{region 'Documentation'}
(*!
<summary>Selects explicit stimuli and expected outcomes; named constants identify every checkpoint.</summary>
*)
{endregion}
METHOD PRIVATE SelectStep : BOOL //! TRUE after selecting a supported script step and its literal expectations; FALSE reports an unknown step.
SelectStep := FALSE;
FRisingFindingExpected := FALSE;
FFallingFindingExpected := FALSE;
FDelayedRisingFindingExpected := FALSE;
FDelayedFallingFindingExpected := FALSE;
CASE FStep OF
    StepInitialBoundReset:
        FTrace := TraceResetHistory;
        FSample := TRUE;
        FSubjectEnable := TRUE;
        FResetSubjects := TRUE;
        FExpectedResult := E_Result.NotEvaluated;
        FExpectedDelayedResult := E_Result.NotEvaluated;
        FExpectedObservation := FALSE;
        FExpectedDelayedObservation := FALSE;
        FExpectedEvaluation := FALSE;
        FExpectedDelayedEvaluation := FALSE;
    StepFirstHighSample:
        FTrace := TraceFirstObservation;
        FSample := TRUE;
        FSubjectEnable := TRUE;
        FResetSubjects := FALSE;
        FExpectedResult := E_Result.NotEvaluated;
        FExpectedDelayedResult := E_Result.NotEvaluated;
        FExpectedObservation := TRUE;
        FExpectedDelayedObservation := FALSE;
        FExpectedEvaluation := FALSE;
        FExpectedDelayedEvaluation := FALSE;
    StepSameHighSample:
        FTrace := TraceFirstObservation;
        FSample := TRUE;
        FSubjectEnable := TRUE;
        FResetSubjects := FALSE;
        FExpectedResult := E_Result.Passed;
        FExpectedDelayedResult := E_Result.NotEvaluated;
        FExpectedObservation := TRUE;
        FExpectedDelayedObservation := TRUE;
        FExpectedEvaluation := TRUE;
        FExpectedDelayedEvaluation := FALSE;
    StepOppositeEdgeAllowed:
        FTrace := TraceFirstObservation;
        FSample := FALSE;
        FSubjectEnable := TRUE;
        FResetSubjects := FALSE;
        FExpectedResult := E_Result.Passed;
        FExpectedDelayedResult := E_Result.Passed;
        FExpectedObservation := TRUE;
        FExpectedDelayedObservation := TRUE;
        FExpectedEvaluation := TRUE;
        FExpectedDelayedEvaluation := TRUE;
    StepForbiddenEdge:
        FTrace := TraceHeldFailure;
        FSample := TRUE;
        FSubjectEnable := TRUE;
        FResetSubjects := FALSE;
        FExpectedResult := E_Result.Failed;
        FExpectedDelayedResult := E_Result.Failed;
        FExpectedObservation := TRUE;
        FExpectedDelayedObservation := TRUE;
        FExpectedEvaluation := TRUE;
        FExpectedDelayedEvaluation := TRUE;
        FRisingFindingExpected := TRUE;
        FFallingFindingExpected := TRUE;
        FDelayedRisingFindingExpected := TRUE;
        FDelayedFallingFindingExpected := TRUE;
    StepRepeatedFailure:
        FTrace := TraceHeldFailure;
        FSample := TRUE;
        FSubjectEnable := TRUE;
        FResetSubjects := FALSE;
        FExpectedResult := E_Result.Failed;
        FExpectedDelayedResult := E_Result.Failed;
        FExpectedObservation := TRUE;
        FExpectedDelayedObservation := TRUE;
        FExpectedEvaluation := TRUE;
        FExpectedDelayedEvaluation := TRUE;
    StepResetBeforeGap:
        FTrace := TraceResetHistory;
        FSample := FALSE;
        FSubjectEnable := TRUE;
        FResetSubjects := TRUE;
        FExpectedResult := E_Result.NotEvaluated;
        FExpectedDelayedResult := E_Result.NotEvaluated;
        FExpectedObservation := FALSE;
        FExpectedDelayedObservation := FALSE;
        FExpectedEvaluation := FALSE;
        FExpectedDelayedEvaluation := FALSE;
    StepBaselineBeforeGap:
        FTrace := TraceDisabledHistory;
        FSample := FALSE;
        FSubjectEnable := TRUE;
        FResetSubjects := FALSE;
        FExpectedResult := E_Result.NotEvaluated;
        FExpectedDelayedResult := E_Result.NotEvaluated;
        FExpectedObservation := TRUE;
        FExpectedDelayedObservation := FALSE;
        FExpectedEvaluation := FALSE;
        FExpectedDelayedEvaluation := FALSE;
    StepDisabledChange:
        FTrace := TraceDisabledHistory;
        FSample := TRUE;
        FSubjectEnable := FALSE;
        FResetSubjects := FALSE;
        FExpectedResult := E_Result.NotEvaluated;
        FExpectedDelayedResult := E_Result.NotEvaluated;
        FExpectedObservation := FALSE;
        FExpectedDelayedObservation := FALSE;
        FExpectedEvaluation := FALSE;
        FExpectedDelayedEvaluation := FALSE;
    StepFirstAfterGap:
        FTrace := TraceDisabledHistory;
        FSample := TRUE;
        FSubjectEnable := TRUE;
        FResetSubjects := FALSE;
        FExpectedResult := E_Result.NotEvaluated;
        FExpectedDelayedResult := E_Result.NotEvaluated;
        FExpectedObservation := TRUE;
        FExpectedDelayedObservation := FALSE;
        FExpectedEvaluation := FALSE;
        FExpectedDelayedEvaluation := FALSE;
    StepSecondAfterGap:
        FTrace := TraceDisabledHistory;
        FSample := TRUE;
        FSubjectEnable := TRUE;
        FResetSubjects := FALSE;
        FExpectedResult := E_Result.Passed;
        FExpectedDelayedResult := E_Result.NotEvaluated;
        FExpectedObservation := TRUE;
        FExpectedDelayedObservation := TRUE;
        FExpectedEvaluation := TRUE;
        FExpectedDelayedEvaluation := FALSE;
    StepAllowedAfterGap:
        FTrace := TraceDisabledHistory;
        FSample := FALSE;
        FSubjectEnable := TRUE;
        FResetSubjects := FALSE;
        FExpectedResult := E_Result.Passed;
        FExpectedDelayedResult := E_Result.Passed;
        FExpectedObservation := TRUE;
        FExpectedDelayedObservation := TRUE;
        FExpectedEvaluation := TRUE;
        FExpectedDelayedEvaluation := TRUE;
    StepForbiddenAfterGap:
        FTrace := TraceDisabledHistory;
        FSample := TRUE;
        FSubjectEnable := TRUE;
        FResetSubjects := FALSE;
        FExpectedResult := E_Result.Failed;
        FExpectedDelayedResult := E_Result.Failed;
        FExpectedObservation := TRUE;
        FExpectedDelayedObservation := TRUE;
        FExpectedEvaluation := TRUE;
        FExpectedDelayedEvaluation := TRUE;
        FRisingFindingExpected := TRUE;
        FFallingFindingExpected := TRUE;
        FDelayedRisingFindingExpected := TRUE;
        FDelayedFallingFindingExpected := TRUE;
    StepResetBeforeDelay:
        FTrace := TraceResetHistory;
        FSample := FALSE;
        FSubjectEnable := TRUE;
        FResetSubjects := TRUE;
        FExpectedResult := E_Result.NotEvaluated;
        FExpectedDelayedResult := E_Result.NotEvaluated;
        FExpectedObservation := FALSE;
        FExpectedDelayedObservation := FALSE;
        FExpectedEvaluation := FALSE;
        FExpectedDelayedEvaluation := FALSE;
    StepSkippedFirstBaseline:
        FTrace := TraceDelayedObservation;
        FSample := FALSE;
        FSubjectEnable := TRUE;
        FResetSubjects := FALSE;
        FExpectedResult := E_Result.NotEvaluated;
        FExpectedDelayedResult := E_Result.NotEvaluated;
        FExpectedObservation := TRUE;
        FExpectedDelayedObservation := FALSE;
        FExpectedEvaluation := FALSE;
        FExpectedDelayedEvaluation := FALSE;
    StepEdgeBeforeDelayedBaseline:
        FTrace := TraceDelayedObservation;
        FSample := TRUE;
        FSubjectEnable := TRUE;
        FResetSubjects := FALSE;
        FExpectedResult := E_Result.Failed;
        FExpectedDelayedResult := E_Result.NotEvaluated;
        FExpectedObservation := TRUE;
        FExpectedDelayedObservation := TRUE;
        FExpectedEvaluation := TRUE;
        FExpectedDelayedEvaluation := FALSE;
        FRisingFindingExpected := TRUE;
        FFallingFindingExpected := TRUE;
    StepStableDelayedBaseline:
        FTrace := TraceDelayedObservation;
        FSample := TRUE;
        FSubjectEnable := TRUE;
        FResetSubjects := FALSE;
        FExpectedResult := E_Result.Failed;
        FExpectedDelayedResult := E_Result.Passed;
        FExpectedObservation := TRUE;
        FExpectedDelayedObservation := TRUE;
        FExpectedEvaluation := TRUE;
        FExpectedDelayedEvaluation := TRUE;
ELSE
    Error(Message := 'Unknown observation trace step.');
    RETURN;
END_CASE;
SelectStep := TRUE;
END_METHOD

END_FUNCTION_BLOCK

// ---- SelfTests/TestCases/TestSuite_AssertionObservation/Test_AssertionEdgeCount.TcPOU
{region 'Documentation'}
(*!
<summary>Checks accumulated rising/falling counts and independent evaluation timing.</summary>
<description>
Both directions run with normal and delayed first observation. Counts survive disabled intervals, but transitions across a gap do not count. Combined observation/evaluation includes the current edge; Evaluate alone observes no edge. Literal counts test the shared algorithm without repeating the comparison operator matrix.
ProcessTests executes one named step per PLC cycle. ProcessAssertions checks that
step before the next call advances it. Every trace has its own outer Assertion;
FirstFailedStep retains the first mismatching checkpoint for online diagnosis.
Expected findings are captured locally and checked before the next step clears
that capture. Subjects are deliberately not called between scripted steps.
</description>
*)
{endregion}
FUNCTION_BLOCK Test_AssertionEdgeCount EXTENDS TestCaseBase
VAR
    FRising : AssertRisingEdgeCntEqual;
    FFalling : AssertFallingEdgeCntEqual;
    FDelayedRising : AssertRisingEdgeCntEqual;
    FDelayedFalling : AssertFallingEdgeCntEqual;
    FCapture : EventBuffer;
    FEvents : ARRAY[1..CaptureLength] OF ST_Event;
    FCaptureFifo : ST_FifoStatus;
    FCaptureStatus : ST_EventBufferStatus;
    FSetupValid : BOOL;
    FStep : UINT;
    FTrace : UINT;
    FFirstFailedStep : UINT;
    FChecked : BOOL;
    FObservationReady : BOOL;
    FStepMatches : BOOL;
    FResultsMatch : BOOL;
    FActivityMatches : BOOL;
    FFindingsMatch : BOOL;
    FCountsMatch : BOOL;
    FSample : BOOL;
    FSubjectEnable : BOOL;
    FSubjectEvaluate : BOOL;
    FResetSubjects : BOOL;
    FExpectedResult : E_Result;
    FExpectedDelayedResult : E_Result;
    FExpectedObservation : BOOL;
    FExpectedDelayedObservation : BOOL;
    FExpectedEvaluation : BOOL;
    FExpectedDelayedEvaluation : BOOL;
    FCountTarget : UINT;
    FExpectedCount : UINT;
    FRisingFindingExpected : BOOL;
    FFallingFindingExpected : BOOL;
    FDelayedRisingFindingExpected : BOOL;
    FDelayedFallingFindingExpected : BOOL;
END_VAR
VAR
    FResetHistory : AssertTrue;
    FCounting : AssertTrue;
    FDisabledHistory : AssertTrue;
    FEvaluationTiming : AssertTrue;
    FWrongCount : AssertTrue;
END_VAR
VAR CONSTANT
    CaptureLength : UINT := 8;
    StepInitialBoundReset : UINT := 1;
    StepFirstBaseline : UINT := 2;
    StepRepeatedBaseline : UINT := 3;
    StepFirstEdge : UINT := 4;
    StepHeldSignal : UINT := 5;
    StepOppositeEdge : UINT := 6;
    StepSecondEdge : UINT := 7;
    StepDisabledChange : UINT := 8;
    StepFirstAfterGap : UINT := 9;
    StepSecondAfterGap : UINT := 10;
    StepOppositeAfterGap : UINT := 11;
    StepThirdEdge : UINT := 12;
    StepEvaluateOnly : UINT := 13;
    StepBaselineBeforeCombined : UINT := 14;
    StepLowBeforeCombined : UINT := 15;
    StepCountBeforeEvaluate : UINT := 16;
    StepResetAfterPass : UINT := 17;
    StepEvaluateOnFirstEnable : UINT := 18;
    StepNewLowBaseline : UINT := 19;
    StepWrongCountFinding : UINT := 20;
    StepWrongCountHeld : UINT := 21;
    StepResetAfterFailure : UINT := 22;
    LastStep : UINT := StepResetAfterFailure;
    TraceResetHistory : UINT := 1;
    TraceCounting : UINT := 2;
    TraceDisabledHistory : UINT := 3;
    TraceEvaluationTiming : UINT := 4;
    TraceWrongCount : UINT := 5;
END_VAR

SUPER^();

{region 'Documentation'}
(*!
<summary>Collects the outer trace checks, never subject results.</summary>
*)
{endregion}
METHOD PROTECTED AggregateResults
VAR_INPUT
    Aggregator : I_ResultAggregator; //! Borrowed result sink owned by the outer Test Case; add this test's checking Assertions without resetting or retaining the sink.
END_VAR
Aggregator.AddProvider(Provider := FResetHistory);
Aggregator.AddProvider(Provider := FCounting);
Aggregator.AddProvider(Provider := FDisabledHistory);
Aggregator.AddProvider(Provider := FEvaluationTiming);
Aggregator.AddProvider(Provider := FWrongCount);
END_METHOD

{region 'Documentation'}
(*!
<summary>Calls each real production subject once with this step's bound inputs.</summary>
*)
{endregion}
METHOD PRIVATE CallSubjects
FRising(Enable := FSubjectEnable,
    Evaluate := FSubjectEvaluate,
    State := E_State.Running,
    IN := FSample,
    Expected := FCountTarget);
FFalling(Enable := FSubjectEnable,
    Evaluate := FSubjectEvaluate,
    State := E_State.Running,
    IN := NOT FSample,
    Expected := FCountTarget);
FDelayedRising(Enable := FSubjectEnable,
    Evaluate := FSubjectEvaluate,
    State := E_State.Running,
    IN := FSample,
    Expected := FCountTarget);
FDelayedFalling(Enable := FSubjectEnable,
    Evaluate := FSubjectEvaluate,
    State := E_State.Running,
    IN := NOT FSample,
    Expected := FCountTarget);
END_METHOD

{region 'Documentation'}
(*!
<summary>Checks per-step finding order, identity and count without retaining old events.</summary>
*)
{endregion}
METHOD PRIVATE CheckFindings
VAR
    Index : UINT;
    FindingMatches : BOOL;
END_VAR
Index := 1;
FFindingsMatch := TRUE;
IF FRisingFindingExpected THEN
    FindingMatches := IsFindingValid(Index := Index,
        ExpectedName := FRising.Name);
    FFindingsMatch := FFindingsMatch AND FindingMatches;
    Index := Index + 1;
END_IF;
IF FFallingFindingExpected THEN
    FindingMatches := IsFindingValid(Index := Index,
        ExpectedName := FFalling.Name);
    FFindingsMatch := FFindingsMatch AND FindingMatches;
    Index := Index + 1;
END_IF;
IF FDelayedRisingFindingExpected THEN
    FindingMatches := IsFindingValid(Index := Index,
        ExpectedName := FDelayedRising.Name);
    FFindingsMatch := FFindingsMatch AND FindingMatches;
    Index := Index + 1;
END_IF;
IF FDelayedFallingFindingExpected THEN
    FindingMatches := IsFindingValid(Index := Index,
        ExpectedName := FDelayedFalling.Name);
    FFindingsMatch := FFindingsMatch AND FindingMatches;
    Index := Index + 1;
END_IF;
FFindingsMatch := FFindingsMatch
    AND (FCaptureStatus.SequenceId = UINT_TO_UDINT(Index - 1))
    AND (FCaptureStatus.LostEventCount = 0);
END_METHOD

{region 'Documentation'}
(*!
<summary>Rejects incomplete local capture, subject or checking-Assertion setup.</summary>
*)
{endregion}
METHOD PROTECTED CheckInitialization : BOOL //! TRUE when the inherited initialization check and this concrete fixture check both accept the setup.
CheckInitialization := SUPER^.CheckInitialization();
IF NOT CheckInitialization THEN
    RETURN;
END_IF;

CheckInitialization := FSetupValid
    AND FResetHistory.IsInitialized
    AND FCounting.IsInitialized
    AND FDisabledHistory.IsInitialized
    AND FEvaluationTiming.IsInitialized
    AND FWrongCount.IsInitialized;
IF NOT CheckInitialization THEN
    EventPublisher.PublishEvent(Event := CreateFrameworkEvent(Name := Name,
        ResourceName := '',
        State := State,
        Severity := E_EventSeverity.Error,
        Message := 'Observation selftest setup failed.'));
END_IF;
END_METHOD

{region 'Documentation'}
(*!
<summary>Compares public results and activity gates against literal step expectations.</summary>
*)
{endregion}
METHOD PRIVATE CheckResults
FResultsMatch := (FRising.Result = FExpectedResult)
    AND (FFalling.Result = FExpectedResult)
    AND (FDelayedRising.Result = FExpectedDelayedResult)
    AND (FDelayedFalling.Result = FExpectedDelayedResult);
FActivityMatches := (FRising.Enabled = FSubjectEnable)
    AND (FRising.ObservationActive = FExpectedObservation)
    AND (FRising.EvaluationActive = FExpectedEvaluation)
    AND (FFalling.Enabled = FSubjectEnable)
    AND (FFalling.ObservationActive = FExpectedObservation)
    AND (FFalling.EvaluationActive = FExpectedEvaluation)
    AND (FDelayedRising.Enabled = FSubjectEnable)
    AND (FDelayedRising.ObservationActive = FExpectedDelayedObservation)
    AND (FDelayedRising.EvaluationActive = FExpectedDelayedEvaluation)
    AND (FDelayedFalling.Enabled = FSubjectEnable)
    AND (FDelayedFalling.ObservationActive = FExpectedDelayedObservation)
    AND (FDelayedFalling.EvaluationActive = FExpectedDelayedEvaluation);
FCountsMatch := (FRising.EdgeCount = FExpectedCount)
    AND (FFalling.EdgeCount = FExpectedCount)
    AND (FDelayedRising.EdgeCount = FExpectedCount)
    AND (FDelayedFalling.EdgeCount = FExpectedCount);
END_METHOD

{region 'Documentation'}
(*!
<summary>Binds isolated subjects and initializes the outer trace Assertions.</summary>
*)
{endregion}
METHOD PROTECTED Configure
VAR
    Initialized : BOOL;
END_VAR
FPreparationStateCount := 0;
FTestStateCount := 1;
FResetHistory.Initialize(Parent := THIS^,
    AssertionName := 'ResetHistory');
FCounting.Initialize(Parent := THIS^,
    AssertionName := 'Counting');
FDisabledHistory.Initialize(Parent := THIS^,
    AssertionName := 'DisabledHistory');
FEvaluationTiming.Initialize(Parent := THIS^,
    AssertionName := 'EvaluationTiming');
FWrongCount.Initialize(Parent := THIS^,
    AssertionName := 'WrongCount');
FSetupValid := FCapture.Initialize(Buffer := FEvents,
    FifoControl := FCaptureFifo,
    Status := FCaptureStatus);
FRising.BindPublisher(Publisher := FCapture);
Initialized := FRising.Initialize(Parent := THIS^,
    AssertionName := 'Rising',
    ObserveFirstCycle := TRUE);
FSetupValid := FSetupValid AND Initialized;
FFalling.BindPublisher(Publisher := FCapture);
Initialized := FFalling.Initialize(Parent := THIS^,
    AssertionName := 'Falling',
    ObserveFirstCycle := TRUE);
FSetupValid := FSetupValid AND Initialized;
FDelayedRising.BindPublisher(Publisher := FCapture);
Initialized := FDelayedRising.Initialize(Parent := THIS^,
    AssertionName := 'DelayedRising',
    ObserveFirstCycle := FALSE);
FSetupValid := FSetupValid AND Initialized;
FDelayedFalling.BindPublisher(Publisher := FCapture);
Initialized := FDelayedFalling.Initialize(Parent := THIS^,
    AssertionName := 'DelayedFalling',
    ObserveFirstCycle := FALSE);
FSetupValid := FSetupValid AND Initialized;
END_METHOD

{region 'Documentation'}
(*!
<summary>Checks one expected local Failed finding; index is bounded by four subjects.</summary>
*)
{endregion}
METHOD PRIVATE IsFindingValid : BOOL //! TRUE when the selected captured finding satisfies the scenario metadata and diagnostic checks.
VAR_INPUT
    Index : UINT; //! One-based index in the retained isolated event capture.
    ExpectedName : STRING(GVL_Constants.NameLength); //! Independently authored Assertion name expected in the selected finding.
END_VAR
IsFindingValid := (FEvents[Index].SequenceId = UINT_TO_UDINT(Index))
    AND (FEvents[Index].Name = ExpectedName)
    AND (FEvents[Index].OwnerScope = E_OwnerScope.Assertion)
    AND (FEvents[Index].EventType = E_EventType.Result)
    AND (FEvents[Index].State = E_State.Running)
    AND (FEvents[Index].Result = E_Result.Failed)
    AND (FEvents[Index].Message <> '');
END_METHOD

{region 'Documentation'}
(*!
<summary>Completes abort; the trace owns no asynchronous resource.</summary>
*)
{endregion}
METHOD PROTECTED ProcessAbort
VAR_INPUT
    Enable : BOOL; //! Phase permission supplied by the owning Test Case; FALSE does not authorize progression, while observation may continue.
END_VAR
IF Enable THEN
    CompleteAbort();
END_IF;
END_METHOD

{region 'Documentation'}
(*!
<summary>Latches the current trace checkpoint before allowing progression.</summary>
*)
{endregion}
METHOD PROTECTED ProcessAssertions
VAR_INPUT
    Enable : BOOL; //! Phase permission supplied by the owning Test Case; FALSE does not authorize progression, while observation may continue.
END_VAR
VAR
    Check : BOOL;
END_VAR
Check := Enable AND FObservationReady;
FResetHistory(Enable := Check AND (FTrace = TraceResetHistory),
    State := State,
    IN := FStepMatches);
FCounting(Enable := Check AND (FTrace = TraceCounting),
    State := State,
    IN := FStepMatches);
FDisabledHistory(Enable := Check AND (FTrace = TraceDisabledHistory),
    State := State,
    IN := FStepMatches);
FEvaluationTiming(Enable := Check AND (FTrace = TraceEvaluationTiming),
    State := State,
    IN := FStepMatches);
FWrongCount(Enable := Check AND (FTrace = TraceWrongCount),
    State := State,
    IN := FStepMatches);
IF Check THEN
    FChecked := TRUE;
END_IF;
END_METHOD

{region 'Documentation'}
(*!
<summary>No Preparation phase is required.</summary>
*)
{endregion}
METHOD PROTECTED ProcessPreparations
VAR_INPUT
    // SA0033: Required hook; this test has no Preparation phase.
    {attribute 'analysis' := '-33'}
    Enable : BOOL; //! Phase permission supplied by the owning Test Case; FALSE does not authorize progression, while observation may continue.
END_VAR
END_METHOD

{region 'Documentation'}
(*!
<summary>Restarts the trace; subjects consume their reset only with bound inputs.</summary>
*)
{endregion}
METHOD PROTECTED ProcessReset
FStep := StepInitialBoundReset;
FTrace := 0;
FFirstFailedStep := 0;
FChecked := FALSE;
FObservationReady := FALSE;
FStepMatches := TRUE;
FResultsMatch := TRUE;
FActivityMatches := TRUE;
FFindingsMatch := TRUE;
FCountsMatch := TRUE;
FCapture.Reset();
ResetSubjects();
FResetHistory.Reset();
FCounting.Reset();
FDisabledHistory.Reset();
FEvaluationTiming.Reset();
FWrongCount.Reset();
CompleteReset();
END_METHOD

{region 'Documentation'}
(*!
<summary>Executes one named step per active cycle, after the previous check was latched.</summary>
*)
{endregion}
METHOD PROTECTED ProcessTests
VAR_INPUT
    Enable : BOOL; //! Phase permission supplied by the owning Test Case; FALSE does not authorize progression, while observation may continue.
END_VAR
IF NOT Enable THEN
    RETURN;
END_IF;

IF FChecked THEN
    FChecked := FALSE;
    FObservationReady := FALSE;
    IF FStep = LastStep THEN
        CompleteTests();
        RETURN;
    END_IF;
    FStep := FStep + 1;
END_IF;

IF NOT SelectStep() THEN
    RETURN;
END_IF;
FCapture.Reset();
IF FResetSubjects THEN
    ResetSubjects();
END_IF;
CallSubjects();
CheckResults();
CheckFindings();
FStepMatches := FResultsMatch AND FActivityMatches AND FFindingsMatch AND FCountsMatch;
IF NOT FStepMatches AND (FFirstFailedStep = 0) THEN
    FFirstFailedStep := FStep;
END_IF;
FObservationReady := TRUE;
END_METHOD

{region 'Documentation'}
(*!
<summary>Queues reset without accessing typed cyclic inputs.</summary>
*)
{endregion}
METHOD PRIVATE ResetSubjects
FRising.Reset();
FFalling.Reset();
FDelayedRising.Reset();
FDelayedFalling.Reset();
END_METHOD

{region 'Documentation'}
(*!
<summary>Selects explicit stimuli and expected outcomes; named constants identify every checkpoint.</summary>
*)
{endregion}
METHOD PRIVATE SelectStep : BOOL //! TRUE after selecting a supported script step and its literal expectations; FALSE reports an unknown step.
SelectStep := FALSE;
FRisingFindingExpected := FALSE;
FFallingFindingExpected := FALSE;
FDelayedRisingFindingExpected := FALSE;
FDelayedFallingFindingExpected := FALSE;
CASE FStep OF
    StepInitialBoundReset:
        FTrace := TraceResetHistory;
        FSample := FALSE;
        FSubjectEnable := TRUE;
        FSubjectEvaluate := FALSE;
        FResetSubjects := TRUE;
        FExpectedResult := E_Result.NotEvaluated;
        FExpectedDelayedResult := E_Result.NotEvaluated;
        FExpectedObservation := FALSE;
        FExpectedDelayedObservation := FALSE;
        FExpectedEvaluation := FALSE;
        FExpectedDelayedEvaluation := FALSE;
        FExpectedCount := 0;
        FCountTarget := 0;
    StepFirstBaseline:
        FTrace := TraceCounting;
        FSample := FALSE;
        FSubjectEnable := TRUE;
        FSubjectEvaluate := FALSE;
        FResetSubjects := FALSE;
        FExpectedResult := E_Result.NotEvaluated;
        FExpectedDelayedResult := E_Result.NotEvaluated;
        FExpectedObservation := TRUE;
        FExpectedDelayedObservation := FALSE;
        FExpectedEvaluation := FALSE;
        FExpectedDelayedEvaluation := FALSE;
        FExpectedCount := 0;
        FCountTarget := 0;
    StepRepeatedBaseline:
        FTrace := TraceCounting;
        FSample := FALSE;
        FSubjectEnable := TRUE;
        FSubjectEvaluate := FALSE;
        FResetSubjects := FALSE;
        FExpectedResult := E_Result.NotEvaluated;
        FExpectedDelayedResult := E_Result.NotEvaluated;
        FExpectedObservation := TRUE;
        FExpectedDelayedObservation := TRUE;
        FExpectedEvaluation := FALSE;
        FExpectedDelayedEvaluation := FALSE;
        FExpectedCount := 0;
        FCountTarget := 0;
    StepFirstEdge:
        FTrace := TraceCounting;
        FSample := TRUE;
        FSubjectEnable := TRUE;
        FSubjectEvaluate := FALSE;
        FResetSubjects := FALSE;
        FExpectedResult := E_Result.NotEvaluated;
        FExpectedDelayedResult := E_Result.NotEvaluated;
        FExpectedObservation := TRUE;
        FExpectedDelayedObservation := TRUE;
        FExpectedEvaluation := FALSE;
        FExpectedDelayedEvaluation := FALSE;
        FExpectedCount := 1;
        FCountTarget := 0;
    StepHeldSignal:
        FTrace := TraceCounting;
        FSample := TRUE;
        FSubjectEnable := TRUE;
        FSubjectEvaluate := FALSE;
        FResetSubjects := FALSE;
        FExpectedResult := E_Result.NotEvaluated;
        FExpectedDelayedResult := E_Result.NotEvaluated;
        FExpectedObservation := TRUE;
        FExpectedDelayedObservation := TRUE;
        FExpectedEvaluation := FALSE;
        FExpectedDelayedEvaluation := FALSE;
        FExpectedCount := 1;
        FCountTarget := 0;
    StepOppositeEdge:
        FTrace := TraceCounting;
        FSample := FALSE;
        FSubjectEnable := TRUE;
        FSubjectEvaluate := FALSE;
        FResetSubjects := FALSE;
        FExpectedResult := E_Result.NotEvaluated;
        FExpectedDelayedResult := E_Result.NotEvaluated;
        FExpectedObservation := TRUE;
        FExpectedDelayedObservation := TRUE;
        FExpectedEvaluation := FALSE;
        FExpectedDelayedEvaluation := FALSE;
        FExpectedCount := 1;
        FCountTarget := 0;
    StepSecondEdge:
        FTrace := TraceCounting;
        FSample := TRUE;
        FSubjectEnable := TRUE;
        FSubjectEvaluate := FALSE;
        FResetSubjects := FALSE;
        FExpectedResult := E_Result.NotEvaluated;
        FExpectedDelayedResult := E_Result.NotEvaluated;
        FExpectedObservation := TRUE;
        FExpectedDelayedObservation := TRUE;
        FExpectedEvaluation := FALSE;
        FExpectedDelayedEvaluation := FALSE;
        FExpectedCount := 2;
        FCountTarget := 0;
    StepDisabledChange:
        FTrace := TraceDisabledHistory;
        FSample := FALSE;
        FSubjectEnable := FALSE;
        FSubjectEvaluate := FALSE;
        FResetSubjects := FALSE;
        FExpectedResult := E_Result.NotEvaluated;
        FExpectedDelayedResult := E_Result.NotEvaluated;
        FExpectedObservation := FALSE;
        FExpectedDelayedObservation := FALSE;
        FExpectedEvaluation := FALSE;
        FExpectedDelayedEvaluation := FALSE;
        FExpectedCount := 2;
        FCountTarget := 0;
    StepFirstAfterGap:
        FTrace := TraceDisabledHistory;
        FSample := TRUE;
        FSubjectEnable := TRUE;
        FSubjectEvaluate := FALSE;
        FResetSubjects := FALSE;
        FExpectedResult := E_Result.NotEvaluated;
        FExpectedDelayedResult := E_Result.NotEvaluated;
        FExpectedObservation := TRUE;
        FExpectedDelayedObservation := FALSE;
        FExpectedEvaluation := FALSE;
        FExpectedDelayedEvaluation := FALSE;
        FExpectedCount := 2;
        FCountTarget := 0;
    StepSecondAfterGap:
        FTrace := TraceDisabledHistory;
        FSample := TRUE;
        FSubjectEnable := TRUE;
        FSubjectEvaluate := FALSE;
        FResetSubjects := FALSE;
        FExpectedResult := E_Result.NotEvaluated;
        FExpectedDelayedResult := E_Result.NotEvaluated;
        FExpectedObservation := TRUE;
        FExpectedDelayedObservation := TRUE;
        FExpectedEvaluation := FALSE;
        FExpectedDelayedEvaluation := FALSE;
        FExpectedCount := 2;
        FCountTarget := 0;
    StepOppositeAfterGap:
        FTrace := TraceDisabledHistory;
        FSample := FALSE;
        FSubjectEnable := TRUE;
        FSubjectEvaluate := FALSE;
        FResetSubjects := FALSE;
        FExpectedResult := E_Result.NotEvaluated;
        FExpectedDelayedResult := E_Result.NotEvaluated;
        FExpectedObservation := TRUE;
        FExpectedDelayedObservation := TRUE;
        FExpectedEvaluation := FALSE;
        FExpectedDelayedEvaluation := FALSE;
        FExpectedCount := 2;
        FCountTarget := 0;
    StepThirdEdge:
        FTrace := TraceDisabledHistory;
        FSample := TRUE;
        FSubjectEnable := TRUE;
        FSubjectEvaluate := FALSE;
        FResetSubjects := FALSE;
        FExpectedResult := E_Result.NotEvaluated;
        FExpectedDelayedResult := E_Result.NotEvaluated;
        FExpectedObservation := TRUE;
        FExpectedDelayedObservation := TRUE;
        FExpectedEvaluation := FALSE;
        FExpectedDelayedEvaluation := FALSE;
        FExpectedCount := 3;
        FCountTarget := 0;
    StepEvaluateOnly:
        FTrace := TraceEvaluationTiming;
        FSample := FALSE;
        FSubjectEnable := FALSE;
        FSubjectEvaluate := TRUE;
        FResetSubjects := FALSE;
        FExpectedResult := E_Result.Passed;
        FExpectedDelayedResult := E_Result.Passed;
        FExpectedObservation := FALSE;
        FExpectedDelayedObservation := FALSE;
        FExpectedEvaluation := TRUE;
        FExpectedDelayedEvaluation := TRUE;
        FExpectedCount := 3;
        FCountTarget := 3;
    StepBaselineBeforeCombined:
        FTrace := TraceEvaluationTiming;
        FSample := TRUE;
        FSubjectEnable := TRUE;
        FSubjectEvaluate := FALSE;
        FResetSubjects := FALSE;
        FExpectedResult := E_Result.Passed;
        FExpectedDelayedResult := E_Result.Passed;
        FExpectedObservation := TRUE;
        FExpectedDelayedObservation := FALSE;
        FExpectedEvaluation := FALSE;
        FExpectedDelayedEvaluation := FALSE;
        FExpectedCount := 3;
        FCountTarget := 0;
    StepLowBeforeCombined:
        FTrace := TraceEvaluationTiming;
        FSample := FALSE;
        FSubjectEnable := TRUE;
        FSubjectEvaluate := FALSE;
        FResetSubjects := FALSE;
        FExpectedResult := E_Result.Passed;
        FExpectedDelayedResult := E_Result.Passed;
        FExpectedObservation := TRUE;
        FExpectedDelayedObservation := TRUE;
        FExpectedEvaluation := FALSE;
        FExpectedDelayedEvaluation := FALSE;
        FExpectedCount := 3;
        FCountTarget := 0;
    StepCountBeforeEvaluate:
        FTrace := TraceEvaluationTiming;
        FSample := TRUE;
        FSubjectEnable := TRUE;
        FSubjectEvaluate := TRUE;
        FResetSubjects := FALSE;
        FExpectedResult := E_Result.Passed;
        FExpectedDelayedResult := E_Result.Passed;
        FExpectedObservation := TRUE;
        FExpectedDelayedObservation := TRUE;
        FExpectedEvaluation := TRUE;
        FExpectedDelayedEvaluation := TRUE;
        FExpectedCount := 4;
        FCountTarget := 4;
    StepResetAfterPass:
        FTrace := TraceResetHistory;
        FSample := TRUE;
        FSubjectEnable := TRUE;
        FSubjectEvaluate := TRUE;
        FResetSubjects := TRUE;
        FExpectedResult := E_Result.NotEvaluated;
        FExpectedDelayedResult := E_Result.NotEvaluated;
        FExpectedObservation := FALSE;
        FExpectedDelayedObservation := FALSE;
        FExpectedEvaluation := FALSE;
        FExpectedDelayedEvaluation := FALSE;
        FExpectedCount := 0;
        FCountTarget := 0;
    StepEvaluateOnFirstEnable:
        FTrace := TraceEvaluationTiming;
        FSample := TRUE;
        FSubjectEnable := TRUE;
        FSubjectEvaluate := TRUE;
        FResetSubjects := FALSE;
        FExpectedResult := E_Result.Passed;
        FExpectedDelayedResult := E_Result.Passed;
        FExpectedObservation := TRUE;
        FExpectedDelayedObservation := FALSE;
        FExpectedEvaluation := TRUE;
        FExpectedDelayedEvaluation := TRUE;
        FExpectedCount := 0;
        FCountTarget := 0;
    StepNewLowBaseline:
        FTrace := TraceWrongCount;
        FSample := FALSE;
        FSubjectEnable := TRUE;
        FSubjectEvaluate := FALSE;
        FResetSubjects := FALSE;
        FExpectedResult := E_Result.Passed;
        FExpectedDelayedResult := E_Result.Passed;
        FExpectedObservation := TRUE;
        FExpectedDelayedObservation := TRUE;
        FExpectedEvaluation := FALSE;
        FExpectedDelayedEvaluation := FALSE;
        FExpectedCount := 0;
        FCountTarget := 0;
    StepWrongCountFinding:
        FTrace := TraceWrongCount;
        FSample := TRUE;
        FSubjectEnable := TRUE;
        FSubjectEvaluate := TRUE;
        FResetSubjects := FALSE;
        FExpectedResult := E_Result.Failed;
        FExpectedDelayedResult := E_Result.Failed;
        FExpectedObservation := TRUE;
        FExpectedDelayedObservation := TRUE;
        FExpectedEvaluation := TRUE;
        FExpectedDelayedEvaluation := TRUE;
        FExpectedCount := 1;
        FCountTarget := 0;
        FRisingFindingExpected := TRUE;
        FFallingFindingExpected := TRUE;
        FDelayedRisingFindingExpected := TRUE;
        FDelayedFallingFindingExpected := TRUE;
    StepWrongCountHeld:
        FTrace := TraceWrongCount;
        FSample := TRUE;
        FSubjectEnable := TRUE;
        FSubjectEvaluate := TRUE;
        FResetSubjects := FALSE;
        FExpectedResult := E_Result.Failed;
        FExpectedDelayedResult := E_Result.Failed;
        FExpectedObservation := TRUE;
        FExpectedDelayedObservation := TRUE;
        FExpectedEvaluation := TRUE;
        FExpectedDelayedEvaluation := TRUE;
        FExpectedCount := 1;
        FCountTarget := 0;
    StepResetAfterFailure:
        FTrace := TraceResetHistory;
        FSample := TRUE;
        FSubjectEnable := TRUE;
        FSubjectEvaluate := TRUE;
        FResetSubjects := TRUE;
        FExpectedResult := E_Result.NotEvaluated;
        FExpectedDelayedResult := E_Result.NotEvaluated;
        FExpectedObservation := FALSE;
        FExpectedDelayedObservation := FALSE;
        FExpectedEvaluation := FALSE;
        FExpectedDelayedEvaluation := FALSE;
        FExpectedCount := 0;
        FCountTarget := 0;
ELSE
    Error(Message := 'Unknown observation trace step.');
    RETURN;
END_CASE;
SelectStep := TRUE;
END_METHOD

END_FUNCTION_BLOCK

// ---- SelfTests/TestCases/TestSuite_AssertionObservation/Test_AssertionSequence.TcPOU
{region 'Documentation'}
(*!
<summary>Checks sequence progress, explicit evaluation, arbitrary lower bounds and deferred reset.</summary>
<description>
DINT Expected starts at -2, BYTE Expected at 4, and a singleton at 8. Expected arrays remain fixed for every run. Reset requests precede the first typed call; only that call binds Expected and consumes reset. Repeated values do not advance, disabled calls retain progress, and explicit Evaluate still checks IN. A separately controlled singleton checks the one-entry boundary.
ProcessTests executes one named step per PLC cycle. ProcessAssertions checks that
step before the next call advances it. Every trace has its own outer Assertion;
FirstFailedStep retains the first mismatching checkpoint for online diagnosis.
Expected findings are captured locally and checked before the next step clears
that capture. Subjects are deliberately not called between scripted steps.
</description>
*)
{endregion}
FUNCTION_BLOCK Test_AssertionSequence EXTENDS TestCaseBase
VAR
    FSequence : AssertSequence_DInt;
    FByteSequence : AssertSequence_Byte;
    FDelayedSequence : AssertSequence_DInt;
    FSingleSequence : AssertSequence_DInt;
    FExpectedSequence : ARRAY[-2..0] OF DINT := [10, 20, 30];
    FExpectedByteSequence : ARRAY[4..6] OF BYTE := [10, 20, 30];
    FExpectedSingle : ARRAY[8..8] OF DINT := [7];
    FCapture : EventBuffer;
    FEvents : ARRAY[1..CaptureLength] OF ST_Event;
    FCaptureFifo : ST_FifoStatus;
    FCaptureStatus : ST_EventBufferStatus;
    FSetupValid : BOOL;
    FStep : UINT;
    FTrace : UINT;
    FFirstFailedStep : UINT;
    FChecked : BOOL;
    FObservationReady : BOOL;
    FStepMatches : BOOL;
    FResultsMatch : BOOL;
    FActivityMatches : BOOL;
    FFindingsMatch : BOOL;
    FSample : DINT;
    FSubjectEnable : BOOL;
    FSubjectEvaluate : BOOL;
    FResetSubjects : BOOL;
    FExpectedResult : E_Result;
    FExpectedDelayedResult : E_Result;
    FExpectedObservation : BOOL;
    FExpectedDelayedObservation : BOOL;
    FExpectedEvaluation : BOOL;
    FExpectedDelayedEvaluation : BOOL;
    FSingleEnable : BOOL;
    FSingleEvaluate : BOOL;
    FSingleSample : DINT;
    FExpectedSingleResult : E_Result;
    FSequenceFindingExpected : BOOL;
    FByteSequenceFindingExpected : BOOL;
    FDelayedSequenceFindingExpected : BOOL;
    FSingleSequenceFindingExpected : BOOL;
END_VAR
VAR
    FDeferredReset : AssertTrue;
    FProgression : AssertTrue;
    FCompletion : AssertTrue;
    FMismatch : AssertTrue;
    FIncomplete : AssertTrue;
    FDisabledProgress : AssertTrue;
    FExplicitEvaluation : AssertTrue;
    FDelayedObservation : AssertTrue;
    FSingleEntry : AssertTrue;
END_VAR
VAR CONSTANT
    CaptureLength : UINT := 8;
    StepInitialBoundReset : UINT := 1;
    StepFirstValue : UINT := 2;
    StepRepeatedFirstValue : UINT := 3;
    StepSecondValue : UINT := 4;
    StepRepeatedSecondValue : UINT := 5;
    StepLastValueWithoutEvaluate : UINT := 6;
    StepEvaluateCompleteDisabled : UINT := 7;
    StepBeyondLastValue : UINT := 8;
    StepBeyondLastAfterDelay : UINT := 9;
    StepResetBeforeMismatch : UINT := 10;
    StepFirstBeforeMismatch : UINT := 11;
    StepRepeatBeforeMismatch : UINT := 12;
    StepSkippedEntry : UINT := 13;
    StepResetBeforeIncomplete : UINT := 14;
    StepFirstBeforeIncomplete : UINT := 15;
    StepRepeatBeforeIncomplete : UINT := 16;
    StepEvaluateIncomplete : UINT := 17;
    StepResetBeforeGap : UINT := 18;
    StepFirstBeforeGap : UINT := 19;
    StepRepeatBeforeGap : UINT := 20;
    StepDisabledUnrelatedValue : UINT := 21;
    StepFirstAfterGap : UINT := 22;
    StepSecondAfterGap : UINT := 23;
    StepCompleteAfterGap : UINT := 24;
    StepResetBeforeEvaluateOnly : UINT := 25;
    StepWrongCurrentValueOnEvaluate : UINT := 26;
    StepResetBeforeFirstCycleEvaluation : UINT := 27;
    StepFirstCycleWrongValue : UINT := 28;
    StepResetBeforeFirstCycleObservation : UINT := 29;
    StepIgnoredFirstCycleValue : UINT := 30;
    StepDelayedFirstValue : UINT := 31;
    StepDelayedSecondValue : UINT := 32;
    StepDelayedCompletion : UINT := 33;
    StepResetBeforeSingleEntry : UINT := 34;
    StepSingleEntryEvaluation : UINT := 35;
    StepSingleEntryContinuation : UINT := 36;
    LastStep : UINT := StepSingleEntryContinuation;
    TraceDeferredReset : UINT := 1;
    TraceProgression : UINT := 2;
    TraceCompletion : UINT := 3;
    TraceMismatch : UINT := 4;
    TraceIncomplete : UINT := 5;
    TraceDisabledProgress : UINT := 6;
    TraceExplicitEvaluation : UINT := 7;
    TraceDelayedObservation : UINT := 8;
    TraceSingleEntry : UINT := 9;
END_VAR

SUPER^();

{region 'Documentation'}
(*!
<summary>Collects the outer trace checks, never subject results.</summary>
*)
{endregion}
METHOD PROTECTED AggregateResults
VAR_INPUT
    Aggregator : I_ResultAggregator; //! Borrowed result sink owned by the outer Test Case; add this test's checking Assertions without resetting or retaining the sink.
END_VAR
Aggregator.AddProvider(Provider := FDeferredReset);
Aggregator.AddProvider(Provider := FProgression);
Aggregator.AddProvider(Provider := FCompletion);
Aggregator.AddProvider(Provider := FMismatch);
Aggregator.AddProvider(Provider := FIncomplete);
Aggregator.AddProvider(Provider := FDisabledProgress);
Aggregator.AddProvider(Provider := FExplicitEvaluation);
Aggregator.AddProvider(Provider := FDelayedObservation);
Aggregator.AddProvider(Provider := FSingleEntry);
END_METHOD

{region 'Documentation'}
(*!
<summary>Calls each real production subject once with this step's bound inputs.</summary>
*)
{endregion}
METHOD PRIVATE CallSubjects
FSequence(Enable := FSubjectEnable,
    Evaluate := FSubjectEvaluate,
    State := E_State.Running,
    IN := FSample,
    Expected := FExpectedSequence);
FByteSequence(Enable := FSubjectEnable,
    Evaluate := FSubjectEvaluate,
    State := E_State.Running,
    IN := DINT_TO_BYTE(FSample),
    Expected := FExpectedByteSequence);
FDelayedSequence(Enable := FSubjectEnable,
    Evaluate := FSubjectEvaluate,
    State := E_State.Running,
    IN := FSample,
    Expected := FExpectedSequence);
FSingleSequence(Enable := FSingleEnable,
    Evaluate := FSingleEvaluate,
    State := E_State.Running,
    IN := FSingleSample,
    Expected := FExpectedSingle);
END_METHOD

{region 'Documentation'}
(*!
<summary>Checks per-step finding order, identity and count without retaining old events.</summary>
*)
{endregion}
METHOD PRIVATE CheckFindings
VAR
    Index : UINT;
    FindingMatches : BOOL;
END_VAR
Index := 1;
FFindingsMatch := TRUE;
IF FSequenceFindingExpected THEN
    FindingMatches := IsFindingValid(Index := Index,
        ExpectedName := FSequence.Name);
    FFindingsMatch := FFindingsMatch AND FindingMatches;
    Index := Index + 1;
END_IF;
IF FByteSequenceFindingExpected THEN
    FindingMatches := IsFindingValid(Index := Index,
        ExpectedName := FByteSequence.Name);
    FFindingsMatch := FFindingsMatch AND FindingMatches;
    Index := Index + 1;
END_IF;
IF FDelayedSequenceFindingExpected THEN
    FindingMatches := IsFindingValid(Index := Index,
        ExpectedName := FDelayedSequence.Name);
    FFindingsMatch := FFindingsMatch AND FindingMatches;
    Index := Index + 1;
END_IF;
IF FSingleSequenceFindingExpected THEN
    FindingMatches := IsFindingValid(Index := Index,
        ExpectedName := FSingleSequence.Name);
    FFindingsMatch := FFindingsMatch AND FindingMatches;
    Index := Index + 1;
END_IF;
FFindingsMatch := FFindingsMatch
    AND (FCaptureStatus.SequenceId = UINT_TO_UDINT(Index - 1))
    AND (FCaptureStatus.LostEventCount = 0);
END_METHOD

{region 'Documentation'}
(*!
<summary>Rejects incomplete local capture, subject or checking-Assertion setup.</summary>
*)
{endregion}
METHOD PROTECTED CheckInitialization : BOOL //! TRUE when the inherited initialization check and this concrete fixture check both accept the setup.
CheckInitialization := SUPER^.CheckInitialization();
IF NOT CheckInitialization THEN
    RETURN;
END_IF;

CheckInitialization := FSetupValid
    AND FDeferredReset.IsInitialized
    AND FProgression.IsInitialized
    AND FCompletion.IsInitialized
    AND FMismatch.IsInitialized
    AND FIncomplete.IsInitialized
    AND FDisabledProgress.IsInitialized
    AND FExplicitEvaluation.IsInitialized
    AND FDelayedObservation.IsInitialized
    AND FSingleEntry.IsInitialized;
IF NOT CheckInitialization THEN
    EventPublisher.PublishEvent(Event := CreateFrameworkEvent(Name := Name,
        ResourceName := '',
        State := State,
        Severity := E_EventSeverity.Error,
        Message := 'Observation selftest setup failed.'));
END_IF;
END_METHOD

{region 'Documentation'}
(*!
<summary>Compares public results and activity gates against literal step expectations.</summary>
*)
{endregion}
METHOD PRIVATE CheckResults
FResultsMatch := (FSequence.Result = FExpectedResult)
    AND (FByteSequence.Result = FExpectedResult)
    AND (FDelayedSequence.Result = FExpectedDelayedResult)
    AND (FSingleSequence.Result = FExpectedSingleResult);
FActivityMatches := (FSequence.Enabled = FSubjectEnable)
    AND (FSequence.ObservationActive = FExpectedObservation)
    AND (FSequence.EvaluationActive = FExpectedEvaluation)
    AND (FByteSequence.Enabled = FSubjectEnable)
    AND (FByteSequence.ObservationActive = FExpectedObservation)
    AND (FByteSequence.EvaluationActive = FExpectedEvaluation)
    AND (FDelayedSequence.Enabled = FSubjectEnable)
    AND (FDelayedSequence.ObservationActive = FExpectedDelayedObservation)
    AND (FDelayedSequence.EvaluationActive = FExpectedDelayedEvaluation)
    AND (FSingleSequence.Enabled = FSingleEnable)
    AND (FSingleSequence.ObservationActive = (FSingleEnable AND NOT FResetSubjects))
    AND (FSingleSequence.EvaluationActive = (FSingleEvaluate AND NOT FResetSubjects));
END_METHOD

{region 'Documentation'}
(*!
<summary>Binds isolated subjects and initializes the outer trace Assertions.</summary>
*)
{endregion}
METHOD PROTECTED Configure
VAR
    Initialized : BOOL;
END_VAR
FPreparationStateCount := 0;
FTestStateCount := 1;
FDeferredReset.Initialize(Parent := THIS^,
    AssertionName := 'DeferredReset');
FProgression.Initialize(Parent := THIS^,
    AssertionName := 'Progression');
FCompletion.Initialize(Parent := THIS^,
    AssertionName := 'Completion');
FMismatch.Initialize(Parent := THIS^,
    AssertionName := 'Mismatch');
FIncomplete.Initialize(Parent := THIS^,
    AssertionName := 'Incomplete');
FDisabledProgress.Initialize(Parent := THIS^,
    AssertionName := 'DisabledProgress');
FExplicitEvaluation.Initialize(Parent := THIS^,
    AssertionName := 'ExplicitEvaluation');
FDelayedObservation.Initialize(Parent := THIS^,
    AssertionName := 'DelayedObservation');
FSingleEntry.Initialize(Parent := THIS^,
    AssertionName := 'SingleEntry');
FSetupValid := FCapture.Initialize(Buffer := FEvents,
    FifoControl := FCaptureFifo,
    Status := FCaptureStatus);
FSequence.BindPublisher(Publisher := FCapture);
Initialized := FSequence.Initialize(Parent := THIS^,
    AssertionName := 'Sequence',
    ObserveFirstCycle := TRUE);
FSetupValid := FSetupValid AND Initialized;
FByteSequence.BindPublisher(Publisher := FCapture);
Initialized := FByteSequence.Initialize(Parent := THIS^,
    AssertionName := 'ByteSequence',
    ObserveFirstCycle := TRUE);
FSetupValid := FSetupValid AND Initialized;
FDelayedSequence.BindPublisher(Publisher := FCapture);
Initialized := FDelayedSequence.Initialize(Parent := THIS^,
    AssertionName := 'DelayedSequence',
    ObserveFirstCycle := FALSE);
FSetupValid := FSetupValid AND Initialized;
FSingleSequence.BindPublisher(Publisher := FCapture);
Initialized := FSingleSequence.Initialize(Parent := THIS^,
    AssertionName := 'SingleSequence',
    ObserveFirstCycle := TRUE);
FSetupValid := FSetupValid AND Initialized;
END_METHOD

{region 'Documentation'}
(*!
<summary>Checks one expected local Failed finding; index is bounded by four subjects.</summary>
*)
{endregion}
METHOD PRIVATE IsFindingValid : BOOL //! TRUE when the selected captured finding satisfies the scenario metadata and diagnostic checks.
VAR_INPUT
    Index : UINT; //! One-based index in the retained isolated event capture.
    ExpectedName : STRING(GVL_Constants.NameLength); //! Independently authored Assertion name expected in the selected finding.
END_VAR
IsFindingValid := (FEvents[Index].SequenceId = UINT_TO_UDINT(Index))
    AND (FEvents[Index].Name = ExpectedName)
    AND (FEvents[Index].OwnerScope = E_OwnerScope.Assertion)
    AND (FEvents[Index].EventType = E_EventType.Result)
    AND (FEvents[Index].State = E_State.Running)
    AND (FEvents[Index].Result = E_Result.Failed)
    AND (FEvents[Index].Message <> '');
END_METHOD

{region 'Documentation'}
(*!
<summary>Completes abort; the trace owns no asynchronous resource.</summary>
*)
{endregion}
METHOD PROTECTED ProcessAbort
VAR_INPUT
    Enable : BOOL; //! Phase permission supplied by the owning Test Case; FALSE does not authorize progression, while observation may continue.
END_VAR
IF Enable THEN
    CompleteAbort();
END_IF;
END_METHOD

{region 'Documentation'}
(*!
<summary>Latches the current trace checkpoint before allowing progression.</summary>
*)
{endregion}
METHOD PROTECTED ProcessAssertions
VAR_INPUT
    Enable : BOOL; //! Phase permission supplied by the owning Test Case; FALSE does not authorize progression, while observation may continue.
END_VAR
VAR
    Check : BOOL;
END_VAR
Check := Enable AND FObservationReady;
FDeferredReset(Enable := Check AND (FTrace = TraceDeferredReset),
    State := State,
    IN := FStepMatches);
FProgression(Enable := Check AND (FTrace = TraceProgression),
    State := State,
    IN := FStepMatches);
FCompletion(Enable := Check AND (FTrace = TraceCompletion),
    State := State,
    IN := FStepMatches);
FMismatch(Enable := Check AND (FTrace = TraceMismatch),
    State := State,
    IN := FStepMatches);
FIncomplete(Enable := Check AND (FTrace = TraceIncomplete),
    State := State,
    IN := FStepMatches);
FDisabledProgress(Enable := Check AND (FTrace = TraceDisabledProgress),
    State := State,
    IN := FStepMatches);
FExplicitEvaluation(Enable := Check AND (FTrace = TraceExplicitEvaluation),
    State := State,
    IN := FStepMatches);
FDelayedObservation(Enable := Check AND (FTrace = TraceDelayedObservation),
    State := State,
    IN := FStepMatches);
FSingleEntry(Enable := Check AND (FTrace = TraceSingleEntry),
    State := State,
    IN := FStepMatches);
IF Check THEN
    FChecked := TRUE;
END_IF;
END_METHOD

{region 'Documentation'}
(*!
<summary>No Preparation phase is required.</summary>
*)
{endregion}
METHOD PROTECTED ProcessPreparations
VAR_INPUT
    // SA0033: Required hook; this test has no Preparation phase.
    {attribute 'analysis' := '-33'}
    Enable : BOOL; //! Phase permission supplied by the owning Test Case; FALSE does not authorize progression, while observation may continue.
END_VAR
END_METHOD

{region 'Documentation'}
(*!
<summary>Restarts the trace; subjects consume their reset only with bound inputs.</summary>
*)
{endregion}
METHOD PROTECTED ProcessReset
FStep := StepInitialBoundReset;
FTrace := 0;
FFirstFailedStep := 0;
FChecked := FALSE;
FObservationReady := FALSE;
FStepMatches := TRUE;
FResultsMatch := TRUE;
FActivityMatches := TRUE;
FFindingsMatch := TRUE;
FCapture.Reset();
ResetSubjects();
FDeferredReset.Reset();
FProgression.Reset();
FCompletion.Reset();
FMismatch.Reset();
FIncomplete.Reset();
FDisabledProgress.Reset();
FExplicitEvaluation.Reset();
FDelayedObservation.Reset();
FSingleEntry.Reset();
CompleteReset();
END_METHOD

{region 'Documentation'}
(*!
<summary>Executes one named step per active cycle, after the previous check was latched.</summary>
*)
{endregion}
METHOD PROTECTED ProcessTests
VAR_INPUT
    Enable : BOOL; //! Phase permission supplied by the owning Test Case; FALSE does not authorize progression, while observation may continue.
END_VAR
IF NOT Enable THEN
    RETURN;
END_IF;

IF FChecked THEN
    FChecked := FALSE;
    FObservationReady := FALSE;
    IF FStep = LastStep THEN
        CompleteTests();
        RETURN;
    END_IF;
    FStep := FStep + 1;
END_IF;

IF NOT SelectStep() THEN
    RETURN;
END_IF;
FCapture.Reset();
IF FResetSubjects THEN
    ResetSubjects();
END_IF;
CallSubjects();
CheckResults();
CheckFindings();
FStepMatches := FResultsMatch AND FActivityMatches AND FFindingsMatch;
IF NOT FStepMatches AND (FFirstFailedStep = 0) THEN
    FFirstFailedStep := FStep;
END_IF;
FObservationReady := TRUE;
END_METHOD

{region 'Documentation'}
(*!
<summary>Queues reset without accessing typed cyclic inputs.</summary>
*)
{endregion}
METHOD PRIVATE ResetSubjects
FSequence.Reset();
FByteSequence.Reset();
FDelayedSequence.Reset();
FSingleSequence.Reset();
END_METHOD

{region 'Documentation'}
(*!
<summary>Selects explicit stimuli and expected outcomes; named constants identify every checkpoint.</summary>
*)
{endregion}
METHOD PRIVATE SelectStep : BOOL //! TRUE after selecting a supported script step and its literal expectations; FALSE reports an unknown step.
SelectStep := FALSE;
FSequenceFindingExpected := FALSE;
FByteSequenceFindingExpected := FALSE;
FDelayedSequenceFindingExpected := FALSE;
FSingleSequenceFindingExpected := FALSE;
FSingleEnable := FALSE;
FSingleEvaluate := FALSE;
FSingleSample := 7;
FExpectedSingleResult := E_Result.NotEvaluated;
CASE FStep OF
    StepInitialBoundReset:
        FTrace := TraceDeferredReset;
        FSample := 10;
        FSubjectEnable := FALSE;
        FSubjectEvaluate := FALSE;
        FResetSubjects := TRUE;
        FExpectedResult := E_Result.NotEvaluated;
        FExpectedDelayedResult := E_Result.NotEvaluated;
        FExpectedObservation := FALSE;
        FExpectedDelayedObservation := FALSE;
        FExpectedEvaluation := FALSE;
        FExpectedDelayedEvaluation := FALSE;
    StepFirstValue:
        FTrace := TraceProgression;
        FSample := 10;
        FSubjectEnable := TRUE;
        FSubjectEvaluate := FALSE;
        FResetSubjects := FALSE;
        FExpectedResult := E_Result.NotEvaluated;
        FExpectedDelayedResult := E_Result.NotEvaluated;
        FExpectedObservation := TRUE;
        FExpectedDelayedObservation := FALSE;
        FExpectedEvaluation := FALSE;
        FExpectedDelayedEvaluation := FALSE;
    StepRepeatedFirstValue:
        FTrace := TraceProgression;
        FSample := 10;
        FSubjectEnable := TRUE;
        FSubjectEvaluate := FALSE;
        FResetSubjects := FALSE;
        FExpectedResult := E_Result.NotEvaluated;
        FExpectedDelayedResult := E_Result.NotEvaluated;
        FExpectedObservation := TRUE;
        FExpectedDelayedObservation := TRUE;
        FExpectedEvaluation := FALSE;
        FExpectedDelayedEvaluation := FALSE;
    StepSecondValue:
        FTrace := TraceProgression;
        FSample := 20;
        FSubjectEnable := TRUE;
        FSubjectEvaluate := FALSE;
        FResetSubjects := FALSE;
        FExpectedResult := E_Result.NotEvaluated;
        FExpectedDelayedResult := E_Result.NotEvaluated;
        FExpectedObservation := TRUE;
        FExpectedDelayedObservation := TRUE;
        FExpectedEvaluation := FALSE;
        FExpectedDelayedEvaluation := FALSE;
    StepRepeatedSecondValue:
        FTrace := TraceProgression;
        FSample := 20;
        FSubjectEnable := TRUE;
        FSubjectEvaluate := FALSE;
        FResetSubjects := FALSE;
        FExpectedResult := E_Result.NotEvaluated;
        FExpectedDelayedResult := E_Result.NotEvaluated;
        FExpectedObservation := TRUE;
        FExpectedDelayedObservation := TRUE;
        FExpectedEvaluation := FALSE;
        FExpectedDelayedEvaluation := FALSE;
    StepLastValueWithoutEvaluate:
        FTrace := TraceProgression;
        FSample := 30;
        FSubjectEnable := TRUE;
        FSubjectEvaluate := FALSE;
        FResetSubjects := FALSE;
        FExpectedResult := E_Result.NotEvaluated;
        FExpectedDelayedResult := E_Result.NotEvaluated;
        FExpectedObservation := TRUE;
        FExpectedDelayedObservation := TRUE;
        FExpectedEvaluation := FALSE;
        FExpectedDelayedEvaluation := FALSE;
    StepEvaluateCompleteDisabled:
        FTrace := TraceCompletion;
        FSample := 30;
        FSubjectEnable := FALSE;
        FSubjectEvaluate := TRUE;
        FResetSubjects := FALSE;
        FExpectedResult := E_Result.Passed;
        FExpectedDelayedResult := E_Result.Passed;
        FExpectedObservation := FALSE;
        FExpectedDelayedObservation := FALSE;
        FExpectedEvaluation := TRUE;
        FExpectedDelayedEvaluation := TRUE;
    StepBeyondLastValue:
        FTrace := TraceCompletion;
        FSample := 40;
        FSubjectEnable := TRUE;
        FSubjectEvaluate := FALSE;
        FResetSubjects := FALSE;
        FExpectedResult := E_Result.Failed;
        FExpectedDelayedResult := E_Result.Passed;
        FExpectedObservation := TRUE;
        FExpectedDelayedObservation := FALSE;
        FExpectedEvaluation := FALSE;
        FExpectedDelayedEvaluation := FALSE;
        FSequenceFindingExpected := TRUE;
        FByteSequenceFindingExpected := TRUE;
    StepBeyondLastAfterDelay:
        FTrace := TraceCompletion;
        FSample := 40;
        FSubjectEnable := TRUE;
        FSubjectEvaluate := FALSE;
        FResetSubjects := FALSE;
        FExpectedResult := E_Result.Failed;
        FExpectedDelayedResult := E_Result.Failed;
        FExpectedObservation := TRUE;
        FExpectedDelayedObservation := TRUE;
        FExpectedEvaluation := FALSE;
        FExpectedDelayedEvaluation := FALSE;
        FDelayedSequenceFindingExpected := TRUE;
    StepResetBeforeMismatch:
        FTrace := TraceDeferredReset;
        FSample := 10;
        FSubjectEnable := FALSE;
        FSubjectEvaluate := FALSE;
        FResetSubjects := TRUE;
        FExpectedResult := E_Result.NotEvaluated;
        FExpectedDelayedResult := E_Result.NotEvaluated;
        FExpectedObservation := FALSE;
        FExpectedDelayedObservation := FALSE;
        FExpectedEvaluation := FALSE;
        FExpectedDelayedEvaluation := FALSE;
    StepFirstBeforeMismatch:
        FTrace := TraceMismatch;
        FSample := 10;
        FSubjectEnable := TRUE;
        FSubjectEvaluate := FALSE;
        FResetSubjects := FALSE;
        FExpectedResult := E_Result.NotEvaluated;
        FExpectedDelayedResult := E_Result.NotEvaluated;
        FExpectedObservation := TRUE;
        FExpectedDelayedObservation := FALSE;
        FExpectedEvaluation := FALSE;
        FExpectedDelayedEvaluation := FALSE;
    StepRepeatBeforeMismatch:
        FTrace := TraceMismatch;
        FSample := 10;
        FSubjectEnable := TRUE;
        FSubjectEvaluate := FALSE;
        FResetSubjects := FALSE;
        FExpectedResult := E_Result.NotEvaluated;
        FExpectedDelayedResult := E_Result.NotEvaluated;
        FExpectedObservation := TRUE;
        FExpectedDelayedObservation := TRUE;
        FExpectedEvaluation := FALSE;
        FExpectedDelayedEvaluation := FALSE;
    StepSkippedEntry:
        FTrace := TraceMismatch;
        FSample := 30;
        FSubjectEnable := TRUE;
        FSubjectEvaluate := FALSE;
        FResetSubjects := FALSE;
        FExpectedResult := E_Result.Failed;
        FExpectedDelayedResult := E_Result.Failed;
        FExpectedObservation := TRUE;
        FExpectedDelayedObservation := TRUE;
        FExpectedEvaluation := FALSE;
        FExpectedDelayedEvaluation := FALSE;
        FSequenceFindingExpected := TRUE;
        FByteSequenceFindingExpected := TRUE;
        FDelayedSequenceFindingExpected := TRUE;
    StepResetBeforeIncomplete:
        FTrace := TraceDeferredReset;
        FSample := 10;
        FSubjectEnable := FALSE;
        FSubjectEvaluate := FALSE;
        FResetSubjects := TRUE;
        FExpectedResult := E_Result.NotEvaluated;
        FExpectedDelayedResult := E_Result.NotEvaluated;
        FExpectedObservation := FALSE;
        FExpectedDelayedObservation := FALSE;
        FExpectedEvaluation := FALSE;
        FExpectedDelayedEvaluation := FALSE;
    StepFirstBeforeIncomplete:
        FTrace := TraceIncomplete;
        FSample := 10;
        FSubjectEnable := TRUE;
        FSubjectEvaluate := FALSE;
        FResetSubjects := FALSE;
        FExpectedResult := E_Result.NotEvaluated;
        FExpectedDelayedResult := E_Result.NotEvaluated;
        FExpectedObservation := TRUE;
        FExpectedDelayedObservation := FALSE;
        FExpectedEvaluation := FALSE;
        FExpectedDelayedEvaluation := FALSE;
    StepRepeatBeforeIncomplete:
        FTrace := TraceIncomplete;
        FSample := 10;
        FSubjectEnable := TRUE;
        FSubjectEvaluate := FALSE;
        FResetSubjects := FALSE;
        FExpectedResult := E_Result.NotEvaluated;
        FExpectedDelayedResult := E_Result.NotEvaluated;
        FExpectedObservation := TRUE;
        FExpectedDelayedObservation := TRUE;
        FExpectedEvaluation := FALSE;
        FExpectedDelayedEvaluation := FALSE;
    StepEvaluateIncomplete:
        FTrace := TraceIncomplete;
        FSample := 20;
        FSubjectEnable := TRUE;
        FSubjectEvaluate := TRUE;
        FResetSubjects := FALSE;
        FExpectedResult := E_Result.Failed;
        FExpectedDelayedResult := E_Result.Failed;
        FExpectedObservation := TRUE;
        FExpectedDelayedObservation := TRUE;
        FExpectedEvaluation := TRUE;
        FExpectedDelayedEvaluation := TRUE;
        FSequenceFindingExpected := TRUE;
        FByteSequenceFindingExpected := TRUE;
        FDelayedSequenceFindingExpected := TRUE;
    StepResetBeforeGap:
        FTrace := TraceDeferredReset;
        FSample := 10;
        FSubjectEnable := FALSE;
        FSubjectEvaluate := FALSE;
        FResetSubjects := TRUE;
        FExpectedResult := E_Result.NotEvaluated;
        FExpectedDelayedResult := E_Result.NotEvaluated;
        FExpectedObservation := FALSE;
        FExpectedDelayedObservation := FALSE;
        FExpectedEvaluation := FALSE;
        FExpectedDelayedEvaluation := FALSE;
    StepFirstBeforeGap:
        FTrace := TraceDisabledProgress;
        FSample := 10;
        FSubjectEnable := TRUE;
        FSubjectEvaluate := FALSE;
        FResetSubjects := FALSE;
        FExpectedResult := E_Result.NotEvaluated;
        FExpectedDelayedResult := E_Result.NotEvaluated;
        FExpectedObservation := TRUE;
        FExpectedDelayedObservation := FALSE;
        FExpectedEvaluation := FALSE;
        FExpectedDelayedEvaluation := FALSE;
    StepRepeatBeforeGap:
        FTrace := TraceDisabledProgress;
        FSample := 10;
        FSubjectEnable := TRUE;
        FSubjectEvaluate := FALSE;
        FResetSubjects := FALSE;
        FExpectedResult := E_Result.NotEvaluated;
        FExpectedDelayedResult := E_Result.NotEvaluated;
        FExpectedObservation := TRUE;
        FExpectedDelayedObservation := TRUE;
        FExpectedEvaluation := FALSE;
        FExpectedDelayedEvaluation := FALSE;
    StepDisabledUnrelatedValue:
        FTrace := TraceDisabledProgress;
        FSample := 99;
        FSubjectEnable := FALSE;
        FSubjectEvaluate := FALSE;
        FResetSubjects := FALSE;
        FExpectedResult := E_Result.NotEvaluated;
        FExpectedDelayedResult := E_Result.NotEvaluated;
        FExpectedObservation := FALSE;
        FExpectedDelayedObservation := FALSE;
        FExpectedEvaluation := FALSE;
        FExpectedDelayedEvaluation := FALSE;
    StepFirstAfterGap:
        FTrace := TraceDisabledProgress;
        FSample := 10;
        FSubjectEnable := TRUE;
        FSubjectEvaluate := FALSE;
        FResetSubjects := FALSE;
        FExpectedResult := E_Result.NotEvaluated;
        FExpectedDelayedResult := E_Result.NotEvaluated;
        FExpectedObservation := TRUE;
        FExpectedDelayedObservation := FALSE;
        FExpectedEvaluation := FALSE;
        FExpectedDelayedEvaluation := FALSE;
    StepSecondAfterGap:
        FTrace := TraceDisabledProgress;
        FSample := 20;
        FSubjectEnable := TRUE;
        FSubjectEvaluate := FALSE;
        FResetSubjects := FALSE;
        FExpectedResult := E_Result.NotEvaluated;
        FExpectedDelayedResult := E_Result.NotEvaluated;
        FExpectedObservation := TRUE;
        FExpectedDelayedObservation := TRUE;
        FExpectedEvaluation := FALSE;
        FExpectedDelayedEvaluation := FALSE;
    StepCompleteAfterGap:
        FTrace := TraceDisabledProgress;
        FSample := 30;
        FSubjectEnable := TRUE;
        FSubjectEvaluate := TRUE;
        FResetSubjects := FALSE;
        FExpectedResult := E_Result.Passed;
        FExpectedDelayedResult := E_Result.Passed;
        FExpectedObservation := TRUE;
        FExpectedDelayedObservation := TRUE;
        FExpectedEvaluation := TRUE;
        FExpectedDelayedEvaluation := TRUE;
    StepResetBeforeEvaluateOnly:
        FTrace := TraceDeferredReset;
        FSample := 10;
        FSubjectEnable := FALSE;
        FSubjectEvaluate := FALSE;
        FResetSubjects := TRUE;
        FExpectedResult := E_Result.NotEvaluated;
        FExpectedDelayedResult := E_Result.NotEvaluated;
        FExpectedObservation := FALSE;
        FExpectedDelayedObservation := FALSE;
        FExpectedEvaluation := FALSE;
        FExpectedDelayedEvaluation := FALSE;
    StepWrongCurrentValueOnEvaluate:
        FTrace := TraceExplicitEvaluation;
        FSample := 30;
        FSubjectEnable := FALSE;
        FSubjectEvaluate := TRUE;
        FResetSubjects := FALSE;
        FExpectedResult := E_Result.Failed;
        FExpectedDelayedResult := E_Result.Failed;
        FExpectedObservation := FALSE;
        FExpectedDelayedObservation := FALSE;
        FExpectedEvaluation := TRUE;
        FExpectedDelayedEvaluation := TRUE;
        FSequenceFindingExpected := TRUE;
        FByteSequenceFindingExpected := TRUE;
        FDelayedSequenceFindingExpected := TRUE;
    StepResetBeforeFirstCycleEvaluation:
        FTrace := TraceDeferredReset;
        FSample := 10;
        FSubjectEnable := FALSE;
        FSubjectEvaluate := FALSE;
        FResetSubjects := TRUE;
        FExpectedResult := E_Result.NotEvaluated;
        FExpectedDelayedResult := E_Result.NotEvaluated;
        FExpectedObservation := FALSE;
        FExpectedDelayedObservation := FALSE;
        FExpectedEvaluation := FALSE;
        FExpectedDelayedEvaluation := FALSE;
    StepFirstCycleWrongValue:
        FTrace := TraceExplicitEvaluation;
        FSample := 99;
        FSubjectEnable := TRUE;
        FSubjectEvaluate := TRUE;
        FResetSubjects := FALSE;
        FExpectedResult := E_Result.Failed;
        FExpectedDelayedResult := E_Result.Failed;
        FExpectedObservation := TRUE;
        FExpectedDelayedObservation := FALSE;
        FExpectedEvaluation := TRUE;
        FExpectedDelayedEvaluation := TRUE;
        FSequenceFindingExpected := TRUE;
        FByteSequenceFindingExpected := TRUE;
        FDelayedSequenceFindingExpected := TRUE;
    StepResetBeforeFirstCycleObservation:
        FTrace := TraceDeferredReset;
        FSample := 10;
        FSubjectEnable := FALSE;
        FSubjectEvaluate := FALSE;
        FResetSubjects := TRUE;
        FExpectedResult := E_Result.NotEvaluated;
        FExpectedDelayedResult := E_Result.NotEvaluated;
        FExpectedObservation := FALSE;
        FExpectedDelayedObservation := FALSE;
        FExpectedEvaluation := FALSE;
        FExpectedDelayedEvaluation := FALSE;
    StepIgnoredFirstCycleValue:
        FTrace := TraceDelayedObservation;
        FSample := 99;
        FSubjectEnable := TRUE;
        FSubjectEvaluate := FALSE;
        FResetSubjects := FALSE;
        FExpectedResult := E_Result.Failed;
        FExpectedDelayedResult := E_Result.NotEvaluated;
        FExpectedObservation := TRUE;
        FExpectedDelayedObservation := FALSE;
        FExpectedEvaluation := FALSE;
        FExpectedDelayedEvaluation := FALSE;
        FSequenceFindingExpected := TRUE;
        FByteSequenceFindingExpected := TRUE;
    StepDelayedFirstValue:
        FTrace := TraceDelayedObservation;
        FSample := 10;
        FSubjectEnable := TRUE;
        FSubjectEvaluate := FALSE;
        FResetSubjects := FALSE;
        FExpectedResult := E_Result.Failed;
        FExpectedDelayedResult := E_Result.NotEvaluated;
        FExpectedObservation := TRUE;
        FExpectedDelayedObservation := TRUE;
        FExpectedEvaluation := FALSE;
        FExpectedDelayedEvaluation := FALSE;
    StepDelayedSecondValue:
        FTrace := TraceDelayedObservation;
        FSample := 20;
        FSubjectEnable := TRUE;
        FSubjectEvaluate := FALSE;
        FResetSubjects := FALSE;
        FExpectedResult := E_Result.Failed;
        FExpectedDelayedResult := E_Result.NotEvaluated;
        FExpectedObservation := TRUE;
        FExpectedDelayedObservation := TRUE;
        FExpectedEvaluation := FALSE;
        FExpectedDelayedEvaluation := FALSE;
    StepDelayedCompletion:
        FTrace := TraceDelayedObservation;
        FSample := 30;
        FSubjectEnable := TRUE;
        FSubjectEvaluate := TRUE;
        FResetSubjects := FALSE;
        FExpectedResult := E_Result.Failed;
        FExpectedDelayedResult := E_Result.Passed;
        FExpectedObservation := TRUE;
        FExpectedDelayedObservation := TRUE;
        FExpectedEvaluation := TRUE;
        FExpectedDelayedEvaluation := TRUE;
    StepResetBeforeSingleEntry:
        FTrace := TraceDeferredReset;
        FSample := 10;
        FSubjectEnable := FALSE;
        FSubjectEvaluate := FALSE;
        FResetSubjects := TRUE;
        FExpectedResult := E_Result.NotEvaluated;
        FExpectedDelayedResult := E_Result.NotEvaluated;
        FExpectedObservation := FALSE;
        FExpectedDelayedObservation := FALSE;
        FExpectedEvaluation := FALSE;
        FExpectedDelayedEvaluation := FALSE;
    StepSingleEntryEvaluation:
        FTrace := TraceSingleEntry;
        FSample := 10;
        FSubjectEnable := FALSE;
        FSubjectEvaluate := FALSE;
        FResetSubjects := FALSE;
        FExpectedResult := E_Result.NotEvaluated;
        FExpectedDelayedResult := E_Result.NotEvaluated;
        FExpectedObservation := FALSE;
        FExpectedDelayedObservation := FALSE;
        FExpectedEvaluation := FALSE;
        FExpectedDelayedEvaluation := FALSE;
        FSingleEnable := TRUE;
        FSingleEvaluate := TRUE;
        FExpectedSingleResult := E_Result.Passed;
    StepSingleEntryContinuation:
        FTrace := TraceSingleEntry;
        FSample := 10;
        FSubjectEnable := FALSE;
        FSubjectEvaluate := FALSE;
        FResetSubjects := FALSE;
        FExpectedResult := E_Result.NotEvaluated;
        FExpectedDelayedResult := E_Result.NotEvaluated;
        FExpectedObservation := FALSE;
        FExpectedDelayedObservation := FALSE;
        FExpectedEvaluation := FALSE;
        FExpectedDelayedEvaluation := FALSE;
        FSingleEnable := TRUE;
        FSingleSample := 8;
        FExpectedSingleResult := E_Result.Failed;
        FSingleSequenceFindingExpected := TRUE;
ELSE
    Error(Message := 'Unknown observation trace step.');
    RETURN;
END_CASE;
SelectStep := TRUE;
END_METHOD

END_FUNCTION_BLOCK

// ---- Framework/Assertions/POU/BasicTypes/DInt/AssertSequence_DInt.TcPOU
{region 'Documentation'}
(*!
<summary>Checks the observed value sequence; Evaluate also checks the current value and
completeness.</summary>
<description>

Uses the whole Expected array from its declared lower bound. Keep its binding, bounds and
values stable until Reset; supply it on reset and disabled FB calls as well.

Observation accepts the current expected value and then permits advancing by one element
on a later change. Repeated equal values do not advance. An unexpected value or an out-of-range
sequence index reports Failed.

Evaluate checks the current value and requires the final expected element to have been
reached; only then can the result become Passed. Disabling observation retains progression.
Reset restarts it.

</description>
*)
{endregion}
FUNCTION_BLOCK AssertSequence_DInt EXTENDS AssertionWithEvaluationBase
VAR_INPUT
    IN : DINT; //! Actual value to observe.
END_VAR
VAR_IN_OUT CONSTANT
    Expected : ARRAY[*] OF DINT; //! Complete expected sequence; read without modifying the supplied array.
END_VAR
VAR
    FExpectedIndex : DINT;
    FSequenceIndexInitialized : BOOL;
    FAllowAdvance : BOOL;
END_VAR

SUPER^();

{region 'Documentation'}
(*!
<summary>Advances at most one entry and checks the current value before explicit completeness evaluation.</summary>
*)
{endregion}
METHOD PROTECTED Assert
VAR
    LowerIndex : DINT;
    UpperIndex : DINT;
    ExpectedValue : DINT;
    MatchesExpected : BOOL;
    AllowAdvance : BOOL;
    Message : STRING(GVL_Constants.MessageLength);
    ExpectedText : STRING(GVL_Constants.AssertionValueLength);
    ActualText : STRING(GVL_Constants.AssertionValueLength);
END_VAR
LowerIndex := LOWER_BOUND(Expected, 1);
UpperIndex := UPPER_BOUND(Expected, 1);

IF NOT FSequenceIndexInitialized THEN
    FExpectedIndex := LowerIndex;
    FSequenceIndexInitialized := TRUE;
END_IF;

IF NOT (ObservationActive OR EvaluationActive) THEN
    RETURN;
END_IF;

IF Result = E_Result.Error THEN
    RETURN;
END_IF;

IF Result = E_Result.Failed THEN
    RETURN;
END_IF;

IF (FExpectedIndex < LowerIndex) OR (FExpectedIndex > UpperIndex) THEN
    Message := CONCAT('Assertion failed: sequence index out of range. ExpectedIndex = ',
        DINT_TO_STRING(FExpectedIndex));
    Message := CONCAT(Message, ', LowerIndex = ');
    Message := CONCAT(Message, DINT_TO_STRING(LowerIndex));
    Message := CONCAT(Message, ', UpperIndex = ');
    Message := CONCAT(Message, DINT_TO_STRING(UpperIndex));
    Message := CONCAT(Message, '.');
    Fail(Message := Message);
    RETURN;
END_IF;

AllowAdvance := FAllowAdvance;
IF ObservationActive THEN
    FAllowAdvance := TRUE;
END_IF;

ExpectedValue := Expected[FExpectedIndex];
MatchesExpected := IN = ExpectedValue;

IF AllowAdvance AND NOT MatchesExpected THEN
    IF FExpectedIndex = UpperIndex THEN
        Message := CONCAT('Assertion failed: sequence continued beyond its last entry. LastIndex = ',
            DINT_TO_STRING(UpperIndex));
        Message := CONCAT(Message, '.');
        Fail(Message := Message);
        RETURN;
    END_IF;

    FExpectedIndex := FExpectedIndex + 1;
    ExpectedValue := Expected[FExpectedIndex];
    MatchesExpected := IN = ExpectedValue;
END_IF;

IF NOT MatchesExpected THEN
    ExpectedText := DINT_TO_STRING(ExpectedValue);
    ActualText := DINT_TO_STRING(IN);
    Message := CONCAT('Assertion failed: sequence value does not match. ExpectedIndex = ',
        DINT_TO_STRING(FExpectedIndex));
    Message := CONCAT(Message, ', Expected = ');
    Message := CONCAT(Message, ExpectedText);
    Message := CONCAT(Message, ', Actual = ');
    Message := CONCAT(Message, ActualText);
    Message := CONCAT(Message, '.');
    Fail(Message := Message);
    RETURN;
END_IF;

IF NOT EvaluationActive THEN
    RETURN;
END_IF;

IF FExpectedIndex <> UpperIndex THEN
    Message := CONCAT('Assertion failed: sequence is incomplete. ExpectedIndex = ',
        DINT_TO_STRING(FExpectedIndex));
    Message := CONCAT(Message, ', LastIndex = ');
    Message := CONCAT(Message, DINT_TO_STRING(UpperIndex));
    Message := CONCAT(Message, '.');
    Fail(Message := Message);
    RETURN;
END_IF;

Pass();
END_METHOD

{region 'Documentation'}
(*!
<summary>Restart progression at the bound Expected array's lower index.</summary>
<description>

Runs only during the reset FB call with Expected supplied, not directly from Reset or
Initialize. Clears permission to advance from a previous observation.

</description>
*)
{endregion}
METHOD PROTECTED ResetAssertion
FExpectedIndex := LOWER_BOUND(Expected, 1);
FSequenceIndexInitialized := TRUE;
FAllowAdvance := FALSE;
END_METHOD

END_FUNCTION_BLOCK

// ---- Framework/Assertions/POU/BasicTypes/Byte/AssertSequence_Byte.TcPOU
{region 'Documentation'}
(*!
<summary>Checks the observed value sequence; Evaluate also checks the current value and
completeness.</summary>
<description>

Uses the whole Expected array from its declared lower bound. Keep its binding, bounds and
values stable until Reset; supply it on reset and disabled FB calls as well.

Observation accepts the current expected value and then permits advancing by one element
on a later change. Repeated equal values do not advance. An unexpected value or an out-of-range
sequence index reports Failed.

Evaluate checks the current value and requires the final expected element to have been
reached; only then can the result become Passed. Disabling observation retains progression.
Reset restarts it.

Mask applies to progression and comparison. An empty mask reports Error.

</description>
*)
{endregion}
FUNCTION_BLOCK AssertSequence_Byte EXTENDS AssertionWithEvaluationBase
VAR_INPUT
    IN : BYTE; //! Actual value to observe.
    Mask : BYTE := 16#FF; //! Bits relevant to sequence progression and comparison.
END_VAR
VAR_IN_OUT CONSTANT
    Expected : ARRAY[*] OF BYTE; //! Complete expected sequence; read without modifying the supplied array.
END_VAR
VAR
    FExpectedIndex : DINT;
    FSequenceIndexInitialized : BOOL;
    FAllowAdvance : BOOL;
END_VAR

SUPER^();

{region 'Documentation'}
(*!
<summary>Advances at most one entry and checks the current value before explicit completeness evaluation.</summary>
*)
{endregion}
METHOD PROTECTED Assert
VAR
    LowerIndex : DINT;
    UpperIndex : DINT;
    ExpectedValue : BYTE;
    MatchesExpected : BOOL;
    AllowAdvance : BOOL;
    Message : STRING(GVL_Constants.MessageLength);
    ExpectedText : STRING(GVL_Constants.AssertionValueLength);
    ActualText : STRING(GVL_Constants.AssertionValueLength);
    MaskText : STRING(GVL_Constants.AssertionValueLength);
END_VAR
VAR CONSTANT
    NoMask : BYTE := 16#00;
    HexDigitCount : USINT := 2;
END_VAR
LowerIndex := LOWER_BOUND(Expected, 1);
UpperIndex := UPPER_BOUND(Expected, 1);

IF NOT FSequenceIndexInitialized THEN
    FExpectedIndex := LowerIndex;
    FSequenceIndexInitialized := TRUE;
END_IF;

IF NOT (ObservationActive OR EvaluationActive) THEN
    RETURN;
END_IF;

IF Result = E_Result.Error THEN
    RETURN;
END_IF;

IF Mask = NoMask THEN
    MaskText := CreateAssertionTextValue_Hex(Value := BYTE_TO_LWORD(Mask),
        DigitCount := HexDigitCount);
    Message := CONCAT('Assertion error: mask must not be empty. Mask = ',
        MaskText);
    Message := CONCAT(Message, '.');
    Error(Message := Message);
    RETURN;
END_IF;

IF Result = E_Result.Failed THEN
    RETURN;
END_IF;

IF (FExpectedIndex < LowerIndex) OR (FExpectedIndex > UpperIndex) THEN
    Message := CONCAT('Assertion failed: sequence index out of range. ExpectedIndex = ',
        DINT_TO_STRING(FExpectedIndex));
    Message := CONCAT(Message, ', LowerIndex = ');
    Message := CONCAT(Message, DINT_TO_STRING(LowerIndex));
    Message := CONCAT(Message, ', UpperIndex = ');
    Message := CONCAT(Message, DINT_TO_STRING(UpperIndex));
    Message := CONCAT(Message, '.');
    Fail(Message := Message);
    RETURN;
END_IF;

AllowAdvance := FAllowAdvance;
IF ObservationActive THEN
    FAllowAdvance := TRUE;
END_IF;

ExpectedValue := Expected[FExpectedIndex];
MatchesExpected := (IN AND Mask) = (ExpectedValue AND Mask);

IF AllowAdvance AND NOT MatchesExpected THEN
    IF FExpectedIndex = UpperIndex THEN
        Message := CONCAT('Assertion failed: sequence continued beyond its last entry. LastIndex = ',
            DINT_TO_STRING(UpperIndex));
        Message := CONCAT(Message, '.');
        Fail(Message := Message);
        RETURN;
    END_IF;

    FExpectedIndex := FExpectedIndex + 1;
    ExpectedValue := Expected[FExpectedIndex];
    MatchesExpected := (IN AND Mask) = (ExpectedValue AND Mask);
END_IF;

IF NOT MatchesExpected THEN
    ExpectedText := CreateAssertionTextValue_Hex(Value := BYTE_TO_LWORD(ExpectedValue),
        DigitCount := HexDigitCount);
    ActualText := CreateAssertionTextValue_Hex(Value := BYTE_TO_LWORD(IN),
        DigitCount := HexDigitCount);
    Message := CONCAT('Assertion failed: sequence value does not match. ExpectedIndex = ',
        DINT_TO_STRING(FExpectedIndex));
    Message := CONCAT(Message, ', Expected = ');
    Message := CONCAT(Message, ExpectedText);
    Message := CONCAT(Message, ', Actual = ');
    Message := CONCAT(Message, ActualText);
    MaskText := CreateAssertionTextValue_Hex(Value := BYTE_TO_LWORD(Mask),
        DigitCount := HexDigitCount);
    Message := CONCAT(Message, ', Mask = ');
    Message := CONCAT(Message, MaskText);
    Message := CONCAT(Message, '.');
    Fail(Message := Message);
    RETURN;
END_IF;

IF NOT EvaluationActive THEN
    RETURN;
END_IF;

IF FExpectedIndex <> UpperIndex THEN
    Message := CONCAT('Assertion failed: sequence is incomplete. ExpectedIndex = ',
        DINT_TO_STRING(FExpectedIndex));
    Message := CONCAT(Message, ', LastIndex = ');
    Message := CONCAT(Message, DINT_TO_STRING(UpperIndex));
    Message := CONCAT(Message, '.');
    Fail(Message := Message);
    RETURN;
END_IF;

Pass();
END_METHOD

{region 'Documentation'}
(*!
<summary>Restart progression at the bound Expected array's lower index.</summary>
<description>

Runs only during the reset FB call with Expected supplied, not directly from Reset or
Initialize. Clears permission to advance from a previous observation.

</description>
*)
{endregion}
METHOD PROTECTED ResetAssertion
FExpectedIndex := LOWER_BOUND(Expected, 1);
FSequenceIndexInitialized := TRUE;
FAllowAdvance := FALSE;
END_METHOD

END_FUNCTION_BLOCK

// ---- SelfTests/TestCases/TestSuite_AssertionObservation/Test_AssertionScalarObservation.TcPOU
{region 'Documentation'}
(*!
<summary>Checks consecutive scalar observations, copied text history and non-finite baselines.</summary>
<description>
DINT, STRING and WSTRING share the finite trace, including a changed mutable text
buffer. REAL/LREAL additionally reject NaN and either infinity on the first active
observation, before a comparison exists. Re-enable replaces scalar observation
history; Reset also clears the held result.
Each named step calls each subject once and checks public gates, result and local
findings before advancing in the next cycle. Outer Assertions collect checkpoints
per trace; subjects never contribute their intentional failures to the test result.
FirstFailedStep retains the first mismatch. No timed stimulus or expected-result
algorithm is used.
</description>
*)
{endregion}
FUNCTION_BLOCK Test_AssertionScalarObservation EXTENDS TestCaseBase
VAR
    FInteger : AssertNoValueChange_DInt;
    FText : AssertNoValueChange_String;
    FWideText : AssertNoValueChange_WString;
    FReal : AssertNoValueChange_Real;
    FLReal : AssertNoValueChange_LReal;
    FSample : DINT;
    FTextSample : STRING(Param_Assertions.AssertionStringLength);
    FWideTextSample : WSTRING(Param_Assertions.AssertionWStringLength);
    FRealSample : AssertionRealRepresentation;
    FLRealSample : AssertionLRealRepresentation;
    FCapture : EventBuffer;
    FEvents : ARRAY[1..CaptureLength] OF ST_Event;
    FCaptureFifo : ST_FifoStatus;
    FCaptureStatus : ST_EventBufferStatus;
    FSetupValid : BOOL;
    FStep : UINT;
    FTrace : UINT;
    FFirstFailedStep : UINT;
    FChecked : BOOL;
    FObservationReady : BOOL;
    FStepMatches : BOOL;
    FResultsMatch : BOOL;
    FActivityMatches : BOOL;
    FFindingsMatch : BOOL;
    FMemoryMatches : BOOL;
    FResetSubjects : BOOL;
    FIntegerEnable : BOOL;
    FIntegerResult : E_Result;
    FIntegerObservation : BOOL;
    FIntegerEvaluation : BOOL;
    FIntegerFinding : E_Result;
    FTextEnable : BOOL;
    FTextResult : E_Result;
    FTextObservation : BOOL;
    FTextEvaluation : BOOL;
    FTextFinding : E_Result;
    FWideTextEnable : BOOL;
    FWideTextResult : E_Result;
    FWideTextObservation : BOOL;
    FWideTextEvaluation : BOOL;
    FWideTextFinding : E_Result;
    FRealEnable : BOOL;
    FRealResult : E_Result;
    FRealObservation : BOOL;
    FRealEvaluation : BOOL;
    FRealFinding : E_Result;
    FLRealEnable : BOOL;
    FLRealResult : E_Result;
    FLRealObservation : BOOL;
    FLRealEvaluation : BOOL;
    FLRealFinding : E_Result;
    FScalarHistory : AssertTrue;
    FReenableBaseline : AssertTrue;
    FResetBaseline : AssertTrue;
    FScalarNonFinite : AssertTrue;
END_VAR
VAR CONSTANT
    CaptureLength : UINT := 8;
    StepInitialReset : UINT := 1;
    StepInitialObservation : UINT := 2;
    StepEqualObservation : UINT := 3;
    StepChangedObservation : UINT := 4;
    StepReturnToInitial : UINT := 5;
    StepReenableReset : UINT := 6;
    StepReenableBaseline : UINT := 7;
    StepBeforeDisable : UINT := 8;
    StepDisabledChange : UINT := 9;
    StepReenabledCapture : UINT := 10;
    StepReenabledComparison : UINT := 11;
    StepResetNewBaseline : UINT := 12;
    StepNewBaselineCapture : UINT := 13;
    StepNewBaselineComparison : UINT := 14;
    StepNaNReset : UINT := 15;
    StepNaNCapture : UINT := 16;
    StepNaNRepeated : UINT := 17;
    StepPositiveInfinityReset : UINT := 18;
    StepPositiveInfinityCapture : UINT := 19;
    StepPositiveInfinityRepeated : UINT := 20;
    StepNegativeInfinityReset : UINT := 21;
    StepNegativeInfinityCapture : UINT := 22;
    StepNegativeInfinityRepeated : UINT := 23;
    LastStep : UINT := StepNegativeInfinityRepeated;
    TraceScalarHistory : UINT := 1;
    TraceReenableBaseline : UINT := 2;
    TraceResetBaseline : UINT := 3;
    TraceScalarNonFinite : UINT := 4;
END_VAR

SUPER^();

{region 'Documentation'}
(*!
<summary>Aggregates only the outer checks, not the intentionally failing subjects.</summary>
*)
{endregion}
METHOD PROTECTED AggregateResults
VAR_INPUT
    Aggregator : I_ResultAggregator; //! Borrowed result sink owned by the outer Test Case; add this test's checking Assertions without resetting or retaining the sink.
END_VAR
Aggregator.AddProvider(Provider := FScalarHistory);
Aggregator.AddProvider(Provider := FReenableBaseline);
Aggregator.AddProvider(Provider := FResetBaseline);
Aggregator.AddProvider(Provider := FScalarNonFinite);
END_METHOD

{region 'Documentation'}
(*!
<summary>Calls each production subject with stable bindings and the selected stimulus.</summary>
*)
{endregion}
METHOD PRIVATE CallSubjects
FInteger(Enable := FIntegerEnable,
    State := E_State.Running,
    IN := FSample);
FText(Enable := FTextEnable,
    State := E_State.Running,
    IN := FTextSample);
FWideText(Enable := FWideTextEnable,
    State := E_State.Running,
    IN := FWideTextSample);
FReal(Enable := FRealEnable,
    State := E_State.Running,
    IN := FRealSample.Value);
FLReal(Enable := FLRealEnable,
    State := E_State.Running,
    IN := FLRealSample.Value);
END_METHOD

{region 'Documentation'}
(*!
<summary>Checks finding order, identities and exact count without retaining prior events.</summary>
*)
{endregion}
METHOD PRIVATE CheckFindings
VAR
    Index : UINT;
    FindingMatches : BOOL;
END_VAR
Index := 1;
FFindingsMatch := TRUE;
IF FIntegerFinding <> E_Result.NotEvaluated THEN
    FindingMatches := IsFindingValid(Index := Index,
        ExpectedName := FInteger.Name,
        ExpectedResult := FIntegerFinding);
    FFindingsMatch := FFindingsMatch AND FindingMatches;
    Index := Index + 1;
END_IF;
IF FTextFinding <> E_Result.NotEvaluated THEN
    FindingMatches := IsFindingValid(Index := Index,
        ExpectedName := FText.Name,
        ExpectedResult := FTextFinding);
    FFindingsMatch := FFindingsMatch AND FindingMatches;
    Index := Index + 1;
END_IF;
IF FWideTextFinding <> E_Result.NotEvaluated THEN
    FindingMatches := IsFindingValid(Index := Index,
        ExpectedName := FWideText.Name,
        ExpectedResult := FWideTextFinding);
    FFindingsMatch := FFindingsMatch AND FindingMatches;
    Index := Index + 1;
END_IF;
IF FRealFinding <> E_Result.NotEvaluated THEN
    FindingMatches := IsFindingValid(Index := Index,
        ExpectedName := FReal.Name,
        ExpectedResult := FRealFinding);
    FFindingsMatch := FFindingsMatch AND FindingMatches;
    Index := Index + 1;
END_IF;
IF FLRealFinding <> E_Result.NotEvaluated THEN
    FindingMatches := IsFindingValid(Index := Index,
        ExpectedName := FLReal.Name,
        ExpectedResult := FLRealFinding);
    FFindingsMatch := FFindingsMatch AND FindingMatches;
    Index := Index + 1;
END_IF;
FFindingsMatch := FFindingsMatch
    AND (FCaptureStatus.SequenceId = UINT_TO_UDINT(Index - 1))
    AND (FCaptureStatus.LostEventCount = 0);
END_METHOD

{region 'Documentation'}
(*!
<summary>Rejects an incomplete capture or subject setup.</summary>
*)
{endregion}
METHOD PROTECTED CheckInitialization : BOOL //! TRUE when the inherited initialization check and this concrete fixture check both accept the setup.
CheckInitialization := SUPER^.CheckInitialization();
IF NOT CheckInitialization THEN
    RETURN;
END_IF;

CheckInitialization := FSetupValid
    AND FScalarHistory.IsInitialized
    AND FReenableBaseline.IsInitialized
    AND FResetBaseline.IsInitialized
    AND FScalarNonFinite.IsInitialized;
IF NOT CheckInitialization THEN
    EventPublisher.PublishEvent(Event := CreateFrameworkEvent(Name := Name,
        ResourceName := '',
        State := State,
        Severity := E_EventSeverity.Error,
        Message := 'Observation selftest setup failed.'));
END_IF;
END_METHOD

{region 'Documentation'}
(*!
<summary>Checks that the read-only mutable text inputs were not modified by observation.</summary>
*)
{endregion}
METHOD PRIVATE CheckMemory
FMemoryMatches := (FTextSample = DINT_TO_STRING(FSample))
    AND (FWideTextSample = DINT_TO_WSTRING(FSample));
END_METHOD

{region 'Documentation'}
(*!
<summary>Checks literal result and observation/evaluation expectations.</summary>
*)
{endregion}
METHOD PRIVATE CheckResults
FResultsMatch := (FInteger.Result = FIntegerResult)
    AND (FText.Result = FTextResult)
    AND (FWideText.Result = FWideTextResult)
    AND (FReal.Result = FRealResult)
    AND (FLReal.Result = FLRealResult);
FActivityMatches := (FInteger.Enabled = FIntegerEnable)
    AND (FInteger.ObservationActive = FIntegerObservation)
    AND (FInteger.EvaluationActive = FIntegerEvaluation)
    AND (FText.Enabled = FTextEnable)
    AND (FText.ObservationActive = FTextObservation)
    AND (FText.EvaluationActive = FTextEvaluation)
    AND (FWideText.Enabled = FWideTextEnable)
    AND (FWideText.ObservationActive = FWideTextObservation)
    AND (FWideText.EvaluationActive = FWideTextEvaluation)
    AND (FReal.Enabled = FRealEnable)
    AND (FReal.ObservationActive = FRealObservation)
    AND (FReal.EvaluationActive = FRealEvaluation)
    AND (FLReal.Enabled = FLRealEnable)
    AND (FLReal.ObservationActive = FLRealObservation)
    AND (FLReal.EvaluationActive = FLRealEvaluation);
END_METHOD

{region 'Documentation'}
(*!
<summary>Initializes outer checks and isolates intentional subject findings.</summary>
*)
{endregion}
METHOD PROTECTED Configure
VAR
    Initialized : BOOL;
END_VAR
FPreparationStateCount := 0;
FTestStateCount := 1;
FScalarHistory.Initialize(Parent := THIS^,
    AssertionName := 'ScalarHistory');
FReenableBaseline.Initialize(Parent := THIS^,
    AssertionName := 'ReenableBaseline');
FResetBaseline.Initialize(Parent := THIS^,
    AssertionName := 'ResetBaseline');
FScalarNonFinite.Initialize(Parent := THIS^,
    AssertionName := 'ScalarNonFinite');
FSetupValid := FCapture.Initialize(Buffer := FEvents,
    FifoControl := FCaptureFifo,
    Status := FCaptureStatus);
FInteger.BindPublisher(Publisher := FCapture);
Initialized := FInteger.Initialize(Parent := THIS^,
    AssertionName := 'Integer',
    ObserveFirstCycle := TRUE);
FSetupValid := FSetupValid AND Initialized;
FText.BindPublisher(Publisher := FCapture);
Initialized := FText.Initialize(Parent := THIS^,
    AssertionName := 'Text',
    ObserveFirstCycle := TRUE);
FSetupValid := FSetupValid AND Initialized;
FWideText.BindPublisher(Publisher := FCapture);
Initialized := FWideText.Initialize(Parent := THIS^,
    AssertionName := 'WideText',
    ObserveFirstCycle := TRUE);
FSetupValid := FSetupValid AND Initialized;
FReal.BindPublisher(Publisher := FCapture);
Initialized := FReal.Initialize(Parent := THIS^,
    AssertionName := 'Real',
    ObserveFirstCycle := TRUE);
FSetupValid := FSetupValid AND Initialized;
FLReal.BindPublisher(Publisher := FCapture);
Initialized := FLReal.Initialize(Parent := THIS^,
    AssertionName := 'LReal',
    ObserveFirstCycle := TRUE);
FSetupValid := FSetupValid AND Initialized;
END_METHOD

{region 'Documentation'}
(*!
<summary>Checks one expected Failed or Error finding from the bounded local capture.</summary>
*)
{endregion}
METHOD PRIVATE IsFindingValid : BOOL //! TRUE when the selected captured finding satisfies the scenario metadata and diagnostic checks.
VAR_INPUT
    Index : UINT; //! One-based index in the retained isolated event capture.
    ExpectedName : STRING(GVL_Constants.NameLength); //! Independently authored Assertion name expected in the selected finding.
    ExpectedResult : E_Result; //! Independently authored finding result.
END_VAR
IsFindingValid := (FEvents[Index].SequenceId = UINT_TO_UDINT(Index))
    AND (FEvents[Index].Name = ExpectedName)
    AND (FEvents[Index].OwnerScope = E_OwnerScope.Assertion)
    AND (FEvents[Index].EventType = E_EventType.Result)
    AND (FEvents[Index].State = E_State.Running)
    AND (FEvents[Index].Result = ExpectedResult)
    AND (FEvents[Index].Message <> '');
END_METHOD

{region 'Documentation'}
(*!
<summary>Completes abort without asynchronous resources.</summary>
*)
{endregion}
METHOD PROTECTED ProcessAbort
VAR_INPUT
    Enable : BOOL; //! Phase permission supplied by the owning Test Case; FALSE does not authorize progression, while observation may continue.
END_VAR
IF Enable THEN
    CompleteAbort();
END_IF;
END_METHOD

{region 'Documentation'}
(*!
<summary>Checks this checkpoint before the next cycle advances the trace.</summary>
*)
{endregion}
METHOD PROTECTED ProcessAssertions
VAR_INPUT
    Enable : BOOL; //! Phase permission supplied by the owning Test Case; FALSE does not authorize progression, while observation may continue.
END_VAR
VAR
    Check : BOOL;
END_VAR
Check := Enable AND FObservationReady;
FScalarHistory(Enable := Check AND (FTrace = TraceScalarHistory),
    State := State,
    IN := FStepMatches);
FReenableBaseline(Enable := Check AND (FTrace = TraceReenableBaseline),
    State := State,
    IN := FStepMatches);
FResetBaseline(Enable := Check AND (FTrace = TraceResetBaseline),
    State := State,
    IN := FStepMatches);
FScalarNonFinite(Enable := Check AND (FTrace = TraceScalarNonFinite),
    State := State,
    IN := FStepMatches);
IF Check THEN
    FChecked := TRUE;
END_IF;
END_METHOD

{region 'Documentation'}
(*!
<summary>No Preparation phase is required.</summary>
*)
{endregion}
METHOD PROTECTED ProcessPreparations
VAR_INPUT
    // SA0033: Required hook; this test has no Preparation phase.
    {attribute 'analysis' := '-33'}
    Enable : BOOL; //! Phase permission supplied by the owning Test Case; FALSE does not authorize progression, while observation may continue.
END_VAR
END_METHOD

{region 'Documentation'}
(*!
<summary>Resets checkpoint bookkeeping and queues each subject reset.</summary>
*)
{endregion}
METHOD PROTECTED ProcessReset
FStep := StepInitialReset;
FTrace := 0;
FFirstFailedStep := 0;
FChecked := FALSE;
FObservationReady := FALSE;
FCapture.Reset();
ResetSubjects();
FScalarHistory.Reset();
FReenableBaseline.Reset();
FResetBaseline.Reset();
FScalarNonFinite.Reset();
CompleteReset();
END_METHOD

{region 'Documentation'}
(*!
<summary>Executes exactly one named checkpoint per active PLC cycle.</summary>
*)
{endregion}
METHOD PROTECTED ProcessTests
VAR_INPUT
    Enable : BOOL; //! Phase permission supplied by the owning Test Case; FALSE does not authorize progression, while observation may continue.
END_VAR
IF NOT Enable THEN
    RETURN;
END_IF;

IF FChecked THEN
    FChecked := FALSE;
    FObservationReady := FALSE;
    IF FStep = LastStep THEN
        CompleteTests();
        RETURN;
    END_IF;
    FStep := FStep + 1;
END_IF;

IF NOT SelectStep() THEN
    RETURN;
END_IF;
FCapture.Reset();
IF FResetSubjects THEN
    ResetSubjects();
END_IF;
CallSubjects();
CheckResults();
CheckMemory();
CheckFindings();
FStepMatches := FResultsMatch AND FActivityMatches AND FMemoryMatches AND FFindingsMatch;
IF NOT FStepMatches AND (FFirstFailedStep = 0) THEN
    FFirstFailedStep := FStep;
END_IF;
FObservationReady := TRUE;
END_METHOD

{region 'Documentation'}
(*!
<summary>Queues subject reset; the next bound call consumes it.</summary>
*)
{endregion}
METHOD PRIVATE ResetSubjects
FInteger.Reset();
FText.Reset();
FWideText.Reset();
FReal.Reset();
FLReal.Reset();
END_METHOD

